// TwinCAT 3 PLC project Untitled2
// ProgramVersion: 3.1.4024.0
// libraries:
//   Tc2_MC2, * (Beckhoff Automation GmbH)
//   Tc2_NC, * (Beckhoff Automation GmbH)
//   Tc2_Standard, * (Beckhoff Automation GmbH)
//   Tc2_System, * (Beckhoff Automation GmbH)
//   Tc3_MC2_AdvancedHoming, * (Beckhoff Automation GmbH)
//   Tc3_Module, * (Beckhoff Automation GmbH)
// project tree:
//   DUTs/ ST_HandoffCmd.TcDUT, ST_HandoffStatus.TcDUT, ST_AxisPlannedReturnCmd.TcDUT, state.TcDUT
//   POUs/ Handoff.TcPOU, ArmCartesian.TcPOU, ArmCartJog.TcPOU, ArmCartJogGen.TcPOU, err.TcPOU, ArmManual.TcPOU, Axis2Sync.TcPOU, handle.TcPOU, InjectorManual.TcPOU, clear_err.TcPOU, init.TcPOU, MAIN.TcPOU, reset.TcPOU, SelfCheck.TcPOU
//   GVLs/ G.TcGVL
//   / PlcTask.TcTTO
// real-time tasks:
//   TASK PlcTask: cycle T#1ms, priority 20, ADS port 350
// motion (NC):
//   TASK NC-Task 1 SAF: cycle T#1ms, priority 4, ADS port 501
//   TASK 1: cycle T#5ms, priority 8, ADS port 511
//   AXIS Axis 1 (id 1)
//     Dynamic: Acceleration=30.3, Deceleration=30.3, Jerk=3060.3
//     Velo: SlowManual=10, FastManual=50, Maximum=30
//     OtherSettings: AllowMotionCmdToSlave=true
//     encoder EncType=19
//       EncPara: ScaleFactorNumerator=2.5, ScaleFactorDenominator=131072, Offset=230, MaxCount=#xffffffff
//     drive DrvType=16
//       DrvPara: MaxCount=#xffffffff, DriveControlDWord=#x00020100
//         Analog: TorqueSetpointScale=10, ScaleFactorActTorque=0.1
//         TimeComp: TaskDelayCycles=1
//     controller CtrType=1
//       CtrPara: PriorControlFactor=1
//         PosDiffControl: Enable=false
//         Observer: BandWidth=20
//   AXIS Axis 2 (id 2)
//     General: UnitName=°
//     Dynamic: Acceleration=10100, Deceleration=10100, Jerk=5100500
//     Velo: SlowManual=1, FastManual=5
//     OtherSettings: AllowMotionCmdToSlave=true
//     encoder EncType=19
//       EncPara: ScaleFactorNumerator=360, ScaleFactorDenominator=131072, Offset=196.397, MaxCount=#xffffffff
//     drive DrvType=16
//       DrvPara: MaxCount=#xffffffff, DriveControlDWord=#x00020000
//         Analog: TorqueSetpointScale=10, ScaleFactorActTorque=0.1
//         TimeComp: TaskDelayCycles=1
//     controller CtrType=1
//       CtrPara: PriorControlFactor=1
//         PosDiffControl: Enable=false
//         Observer: BandWidth=20
//   AXIS Axis 3 (id 3)
//     General: UnitName=°
//     Velo: SlowManual=3, FastManual=10
//     OtherSettings: AllowMotionCmdToSlave=true
//     encoder EncType=19
//       EncPara: ScaleFactorNumerator=360, ScaleFactorDenominator=131072, Offset=480, MaxCount=#xffffffff
//     drive DrvType=16
//       DrvPara: MaxCount=#xffffffff, DriveControlDWord=#x00020000
//         Analog: TorqueSetpointScale=10, ScaleFactorActTorque=0.1
//         TimeComp: TaskDelayCycles=1
//     controller CtrType=1
//       CtrPara: PriorControlFactor=1
//         PosDiffControl: Enable=false
//         Observer: BandWidth=20
//   AXIS Axis 4 (id 4)
//     General: UnitName=°
//     Dynamic: Acceleration=1570, Deceleration=1570, Jerk=2162.19
//     Velo: SlowManual=3, FastManual=10
//     OtherSettings: AllowMotionCmdToSlave=true
//     encoder EncType=19
//       EncPara: ScaleFactorNumerator=360, ScaleFactorDenominator=131072, Offset=54, MaxCount=#xffffffff
//     drive DrvType=16
//       DrvPara: MaxCount=#xffffffff, DriveControlDWord=#x00020000
//         Analog: TorqueSetpointScale=10, ScaleFactorActTorque=0.1
//         TimeComp: TaskDelayCycles=1
//     controller CtrType=1
//       CtrPara: PriorControlFactor=1
//         PosDiffControl: Enable=false
//         Observer: BandWidth=20
//   AXIS Axis 5 (id 5)
//     General: UnitName=°
//     Velo: SlowManual=3, FastManual=10
//     OtherSettings: AllowMotionCmdToSlave=true
//     encoder EncType=19
//       EncPara: ScaleFactorNumerator=360, ScaleFactorDenominator=131072, MaxCount=#xffffffff
//     drive DrvType=16
//       DrvPara: MaxCount=#xffffffff, DriveControlDWord=#x00020000
//         Analog: TorqueSetpointScale=10, ScaleFactorActTorque=0.1
//         TimeComp: TaskDelayCycles=1
//     controller CtrType=1
//       CtrPara: PriorControlFactor=1
//         Observer: BandWidth=20
//   AXIS Axis 6 (id 6)
//     Velo: SlowManual=3, FastManual=10
//     OtherSettings: AllowMotionCmdToSlave=true
//     encoder EncType=19
//       EncPara: ScaleFactorNumerator=65.94, ScaleFactorDenominator=425164.8, MaxCount=#xffffffff
//     drive DrvType=16
//       DrvPara: MaxCount=#xffffffff, DriveControlDWord=#x00020100
//         Analog: TorqueSetpointScale=10, ScaleFactorActTorque=0.1
//         TimeComp: TaskDelayCycles=1
//     controller CtrType=1
//       CtrPara: PriorControlFactor=1
//         PosDiffControl: Enable=false
//         Observer: BandWidth=20
//   AXIS Axis 7 (id 7)
//     Velo: SlowManual=3, FastManual=10
//     OtherSettings: AllowMotionCmdToSlave=true
//     encoder EncType=19
//       EncPara: ScaleFactorNumerator=360, ScaleFactorDenominator=768300, MaxCount=#xffffffff
//     drive DrvType=16
//       DrvPara: MaxCount=#xffffffff, DriveControlDWord=#x00020000
//         Analog: TorqueSetpointScale=10, ScaleFactorActTorque=0.1
//         TimeComp: TaskDelayCycles=1
//     controller CtrType=1
//       CtrPara: PriorControlFactor=1
//         PosDiffControl: Enable=false
//         Observer: BandWidth=20
//   AXIS Axis 8 (id 8)
//     Velo: SlowManual=3, FastManual=10
//     OtherSettings: AllowMotionCmdToSlave=true
//     encoder EncType=19
//       EncPara: ScaleFactorNumerator=65.94, ScaleFactorDenominator=425164.8, MaxCount=#xffffffff
//     drive DrvType=16
//       DrvPara: MaxCount=#xffffffff, DriveControlDWord=#x00020100
//         Analog: TorqueSetpointScale=10, ScaleFactorActTorque=0.1
//         TimeComp: TaskDelayCycles=1
//     controller CtrType=1
//       CtrPara: PriorControlFactor=1
//         PosDiffControl: Enable=false
//         Observer: BandWidth=20
//   AXIS Axis 9 (id 9)
//     Dynamic: Acceleration=1010, Deceleration=1010, Jerk=51005
//     Velo: SlowManual=3, FastManual=10
//     OtherSettings: AllowMotionCmdToSlave=true
//     encoder EncType=19
//       EncPara: ScaleFactorNumerator=360, ScaleFactorDenominator=758988.8, MaxCount=#xffffffff
//     drive DrvType=16
//       DrvPara: MaxCount=#xffffffff, DriveControlDWord=#x00020000
//         Analog: TorqueSetpointScale=10, ScaleFactorActTorque=0.1
//         TimeComp: TaskDelayCycles=1
//     controller CtrType=1
//       CtrPara: PriorControlFactor=1
//         Observer: BandWidth=20
//   AXIS Axis 10 (id 10)
//     Dynamic: Acceleration=2000, Deceleration=2000, Jerk=2000
//     Velo: SlowManual=3, FastManual=10
//     OtherSettings: AllowMotionCmdToSlave=true
//     encoder EncType=19
//       EncPara: ScaleFactorNumerator=65.94, ScaleFactorDenominator=425164.8, MaxCount=#xffffffff
//     drive DrvType=16
//       DrvPara: MaxCount=#xffffffff, DriveControlDWord=#x00020100
//         Analog: TorqueSetpointScale=10, ScaleFactorActTorque=0.1
//         TimeComp: TaskDelayCycles=1
//     controller CtrType=1
//       CtrPara: PriorControlFactor=1
//         PosDiffControl: Enable=false
//         Observer: BandWidth=20
//   AXIS Axis 11 (id 11)
//     Dynamic: Acceleration=375, Deceleration=375, Jerk=5625
//     Velo: SlowManual=3, FastManual=10
//     OtherSettings: AllowMotionCmdToSlave=true
//     encoder EncType=19
//       EncPara: ScaleFactorNumerator=65.94, ScaleFactorDenominator=425164.8, Inverse=true, MaxCount=#xffffffff
//     drive DrvType=16
//       DrvPara: Inverse=true, MaxCount=#xffffffff, DriveControlDWord=#x00020100
//         Analog: TorqueSetpointScale=10, ScaleFactorActTorque=0.1
//         TimeComp: TaskDelayCycles=1
//     controller CtrType=1
//       CtrPara: PriorControlFactor=1
//         PosDiffControl: Enable=false
//         Observer: BandWidth=20
//   AXIS Axis 12 (id 12)
//     Velo: SlowManual=3, FastManual=10
//     OtherSettings: AllowMotionCmdToSlave=true
//     encoder EncType=19
//       EncPara: ScaleFactorNumerator=360, ScaleFactorDenominator=768300, MaxCount=#xffffffff
//     drive DrvType=16
//       DrvPara: MaxCount=#xffffffff, DriveControlDWord=#x00020000
//         Analog: TorqueSetpointScale=10, ScaleFactorActTorque=0.1
//         TimeComp: TaskDelayCycles=1
//     controller CtrType=1
//       CtrPara: PriorControlFactor=1
//         PosDiffControl: Enable=false
//         Observer: BandWidth=20
//   AXIS Axis 13 (id 13)
//     General: UnitName=°
//     Dynamic: Acceleration=10600, Deceleration=10600, Jerk=936333
//     OtherSettings: AllowMotionCmdToSlave=true
//     encoder EncType=19
//       EncPara: ScaleFactorNumerator=360, ScaleFactorDenominator=180224, MaxCount=#xffffffff
//     drive DrvType=16
//       DrvPara: MaxCount=#xffffffff, DriveControlDWord=#x00020100
//         Analog: TorqueSetpointScale=10, ScaleFactorActTorque=0.1
//         TimeComp: TaskDelayCycles=1
//     controller CtrType=1
//       CtrPara: PriorControlFactor=1
//         PosDiffControl: Enable=false
//         Observer: BandWidth=20
//   AXIS Axis 14 (id 14)
//     General: UnitName=°
//     Dynamic: Acceleration=10400, Deceleration=10400, Jerk=1352000
//     OtherSettings: AllowMotionCmdToSlave=true
//     encoder EncType=19
//       EncPara: ScaleFactorNumerator=360, ScaleFactorDenominator=180224, MaxCount=#xffffffff
//     drive DrvType=16
//       DrvPara: MaxCount=#xffffffff, DriveControlDWord=#x00020100
//         Analog: TorqueSetpointScale=10, ScaleFactorActTorque=0.1
//         TimeComp: TaskDelayCycles=1
//     controller CtrType=1
//       CtrPara: PriorControlFactor=1
//         PosDiffControl: Enable=false
//         Observer: BandWidth=20
//   AXIS Axis 15 (id 15)
//     General: UnitName=°
//     Dynamic: Acceleration=11000, Deceleration=11000, Jerk=605000
//     OtherSettings: AllowMotionCmdToSlave=true
//     encoder EncType=19
//       EncPara: ScaleFactorNumerator=360, ScaleFactorDenominator=757760, MaxCount=#xffffffff
//     drive DrvType=16
//       DrvPara: MaxCount=#xffffffff, DriveControlDWord=#x00020100
//         Analog: TorqueSetpointScale=10, ScaleFactorActTorque=0.1
//         TimeComp: TaskDelayCycles=1
//     controller CtrType=1
//       CtrPara: PriorControlFactor=1
//         PosDiffControl: Enable=false
//         Observer: BandWidth=20
// I/O:
//   DEVICE Device 5 (EtherCAT), AmsNetId 169.254.119.135.6.1
//     Box 1 (EtherCat-control-node) [EtherCat-control-V1.6]
//     Drive 2 (Micro 4804 MZ-CAT-STO ) [Micro 4804 MZ-CAT-STO]
//     Drive 3 (TK Drive ) [EtherCAT Drive Rev:0x00010420]
//     Drive 4 (TK Drive ) [EtherCAT Drive Rev:0x00010420]
//     Drive 5 (TK Drive ) [EtherCAT Drive Rev:0x00010420]
//     Drive 6 (TK Drive ) [EtherCAT Drive Rev:0x00010420]
//     Box 7 (EtherCat-control-node) [EtherCat-control-V1.6]
//     Box 8 (EtherCat-control-node) [EtherCat-control-V1.6]
//     Drive 9 (Micro 4804 MZ-CAT-STO ) [Micro 4804 MZ-CAT-STO]
//     Drive 10 (DEN-XCR-E) [DEN-XCR-E]
//     Drive 11 (Micro 4804 MZ-CAT-STO ) [Micro 4804 MZ-CAT-STO]
//     Drive 12 (DEN-XCR-E) [DEN-XCR-E]
//     Drive 13 (Micro 4804 MZ-CAT-STO ) [Micro 4804 MZ-CAT-STO]
//     Drive 14 (Micro 4804 MZ-CAT-STO ) [Micro 4804 MZ-CAT-STO]
//     Drive 15 (CAP-XCR-E) [CAP-XCR-E]
//     Drive 16 (Micro 4804 MZ-CAT-STO ) [Micro 4804 MZ-CAT-STO]
//     Drive 17 (Micro 4804 MZ-CAT-STO ) [Micro 4804 MZ-CAT-STO]
//     Drive 18 (Micro 4804 MZ-CAT-STO ) [Micro 4804 MZ-CAT-STO]
// variable links:
//   NC-Task 1 SAF/Axes/Axis 1 <-> Device 5 (EtherCAT)/Drive 2 (Micro 4804 MZ-CAT-STO )
//     Drive/Inputs/In/nDataIn1 <-> Transmit PDO 2 mapping parameters/Following error actual value
//     Drive/Inputs/In/nDataIn3[0] <-> Transmit PDO 1 mapping parameters/Torque (current) actual value
//     Drive/Inputs/In/nDcOutputTime <-> InfoData/DcOutputShift
//     Drive/Inputs/In/nState1 <-> Transmit PDO 1 mapping parameters/Statusword
//     Drive/Inputs/In/nState2 <-> Transmit PDO 1 mapping parameters/Statusword @bit 8
//     Drive/Inputs/In/nState4 @bit 1 <-> WcState/InputToggle
//     Drive/Inputs/In/nState4 <-> WcState/WcState
//     Drive/Inputs/In/nState5 <-> Transmit PDO 4 mapping parameters/Modes of operation display
//     Drive/Outputs/Out/nCtrl1 <-> Receive PDO 1 mapping parameters/Controlword
//     Drive/Outputs/Out/nCtrl2 <-> Receive PDO 1 mapping parameters/Controlword @bit 8
//     Drive/Outputs/Out/nCtrl5 <-> Receive PDO 3 mapping parameters/Modes of operation
//     Drive/Outputs/Out/nDataOut1 <-> Receive PDO 1 mapping parameters/Target position
//     Drive/Outputs/Out/nDataOut4[0] <-> Receive PDO 3 mapping parameters/Target torque
//     Enc/Inputs/In/nDataIn1 <-> Transmit PDO 1 mapping parameters/Position actual value
//     Enc/Inputs/In/nDataIn7 <-> Transmit PDO 3 mapping parameters/Velocity actual value
//     Enc/Inputs/In/nDcInputTime <-> InfoData/DcInputShift
//     Enc/Inputs/In/nState4 @bit 1 <-> WcState/InputToggle
//     Enc/Inputs/In/nState4 <-> WcState/WcState
//   NC-Task 1 SAF/Axes/Axis 10 <-> Device 5 (EtherCAT)/Drive 13 (Micro 4804 MZ-CAT-STO )
//     Drive/Inputs/In/nDataIn1 <-> Transmit PDO 2 mapping parameters/Following error actual value
//     Drive/Inputs/In/nDataIn3[0] <-> Transmit PDO 1 mapping parameters/Torque (current) actual value
//     Drive/Inputs/In/nDcOutputTime <-> InfoData/DcOutputShift
//     Drive/Inputs/In/nState1 <-> Transmit PDO 1 mapping parameters/Statusword
//     Drive/Inputs/In/nState2 <-> Transmit PDO 1 mapping parameters/Statusword @bit 8
//     Drive/Inputs/In/nState4 @bit 1 <-> WcState/InputToggle
//     Drive/Inputs/In/nState4 <-> WcState/WcState
//     Drive/Outputs/Out/nCtrl1 <-> Receive PDO 1 mapping parameters/Controlword
//     Drive/Outputs/Out/nCtrl2 <-> Receive PDO 1 mapping parameters/Controlword @bit 8
//     Drive/Outputs/Out/nDataOut1 <-> Receive PDO 1 mapping parameters/Target position
//     Enc/Inputs/In/nDataIn1 <-> Transmit PDO 1 mapping parameters/Position actual value
//     Enc/Inputs/In/nDcInputTime <-> InfoData/DcInputShift
//     Enc/Inputs/In/nState4 @bit 1 <-> WcState/InputToggle
//     Enc/Inputs/In/nState4 <-> WcState/WcState
//   NC-Task 1 SAF/Axes/Axis 11 <-> Device 5 (EtherCAT)/Drive 14 (Micro 4804 MZ-CAT-STO )
//     Drive/Inputs/In/nDataIn1 <-> Transmit PDO 2 mapping parameters/Following error actual value
//     Drive/Inputs/In/nDataIn3[0] <-> Transmit PDO 1 mapping parameters/Torque (current) actual value
//     Drive/Inputs/In/nDcOutputTime <-> InfoData/DcOutputShift
//     Drive/Inputs/In/nState1 <-> Transmit PDO 1 mapping parameters/Statusword
//     Drive/Inputs/In/nState2 <-> Transmit PDO 1 mapping parameters/Statusword @bit 8
//     Drive/Inputs/In/nState4 @bit 1 <-> WcState/InputToggle
//     Drive/Inputs/In/nState4 <-> WcState/WcState
//     Drive/Outputs/Out/nCtrl1 <-> Receive PDO 1 mapping parameters/Controlword
//     Drive/Outputs/Out/nCtrl2 <-> Receive PDO 1 mapping parameters/Controlword @bit 8
//     Drive/Outputs/Out/nDataOut1 <-> Receive PDO 1 mapping parameters/Target position
//     Enc/Inputs/In/nDataIn1 <-> Transmit PDO 1 mapping parameters/Position actual value
//     Enc/Inputs/In/nDcInputTime <-> InfoData/DcInputShift
//     Enc/Inputs/In/nState4 @bit 1 <-> WcState/InputToggle
//     Enc/Inputs/In/nState4 <-> WcState/WcState
//   NC-Task 1 SAF/Axes/Axis 12 <-> Device 5 (EtherCAT)/Drive 15 (CAP-XCR-E)
//     Drive/Inputs/In/nState1 <-> TPDO 1 mapping parameter/Status Word
//     Drive/Inputs/In/nState2 <-> TPDO 1 mapping parameter/Status Word @bit 8
//     Drive/Inputs/In/nState4 @bit 1 <-> WcState/InputToggle
//     Drive/Inputs/In/nState4 <-> WcState/WcState
//     Drive/Inputs/In/nState5 <-> TPDO 1 mapping parameter/Operation mode display
//     Drive/Outputs/Out/nCtrl1 <-> RPDO 1 mapping parameter/Control Word
//     Drive/Outputs/Out/nCtrl2 <-> RPDO 1 mapping parameter/Control Word @bit 8
//     Drive/Outputs/Out/nCtrl5 <-> RPDO 1 mapping parameter/Operation mode
//     Drive/Outputs/Out/nDataOut1 <-> RPDO 1 mapping parameter/Position set-point
//     Drive/Outputs/Out/nDataOut2 <-> RPDO 1 mapping parameter/Velocity set-point
//     Enc/Inputs/In/nDataIn1 <-> TPDO 1 mapping parameter/Actual position
//     Enc/Inputs/In/nDataIn7 <-> TPDO 1 mapping parameter/Actual velocity
//     Enc/Inputs/In/nState4 @bit 1 <-> WcState/InputToggle
//     Enc/Inputs/In/nState4 <-> WcState/WcState
//   NC-Task 1 SAF/Axes/Axis 13 <-> Device 5 (EtherCAT)/Drive 16 (Micro 4804 MZ-CAT-STO )
//     Drive/Inputs/In/nDataIn1 <-> Transmit PDO 2 mapping parameters/Following error actual value
//     Drive/Inputs/In/nDataIn3[0] <-> Transmit PDO 1 mapping parameters/Torque (current) actual value
//     Drive/Inputs/In/nDcOutputTime <-> InfoData/DcOutputShift
//     Drive/Inputs/In/nState1 <-> Transmit PDO 1 mapping parameters/Statusword
//     Drive/Inputs/In/nState2 <-> Transmit PDO 1 mapping parameters/Statusword @bit 8
//     Drive/Inputs/In/nState4 @bit 1 <-> WcState/InputToggle
//     Drive/Inputs/In/nState4 <-> WcState/WcState
//     Drive/Outputs/Out/nCtrl1 <-> Receive PDO 1 mapping parameters/Controlword
//     Drive/Outputs/Out/nCtrl2 <-> Receive PDO 1 mapping parameters/Controlword @bit 8
//     Drive/Outputs/Out/nDataOut1 <-> Receive PDO 1 mapping parameters/Target position
//     Enc/Inputs/In/nDataIn1 <-> Transmit PDO 1 mapping parameters/Position actual value
//     Enc/Inputs/In/nDcInputTime <-> InfoData/DcInputShift
//     Enc/Inputs/In/nState4 @bit 1 <-> WcState/InputToggle
//     Enc/Inputs/In/nState4 <-> WcState/WcState
//   NC-Task 1 SAF/Axes/Axis 14 <-> Device 5 (EtherCAT)/Drive 17 (Micro 4804 MZ-CAT-STO )
//     Drive/Inputs/In/nDataIn1 <-> Transmit PDO 2 mapping parameters/Following error actual value
//     Drive/Inputs/In/nDataIn3[0] <-> Transmit PDO 1 mapping parameters/Torque (current) actual value
//     Drive/Inputs/In/nDcOutputTime <-> InfoData/DcOutputShift
//     Drive/Inputs/In/nState1 <-> Transmit PDO 1 mapping parameters/Statusword
//     Drive/Inputs/In/nState2 <-> Transmit PDO 1 mapping parameters/Statusword @bit 8
//     Drive/Inputs/In/nState4 @bit 1 <-> WcState/InputToggle
//     Drive/Inputs/In/nState4 <-> WcState/WcState
//     Drive/Outputs/Out/nCtrl1 <-> Receive PDO 1 mapping parameters/Controlword
//     Drive/Outputs/Out/nCtrl2 <-> Receive PDO 1 mapping parameters/Controlword @bit 8
//     Drive/Outputs/Out/nDataOut1 <-> Receive PDO 1 mapping parameters/Target position
//     Enc/Inputs/In/nDataIn1 <-> Transmit PDO 1 mapping parameters/Position actual value
//     Enc/Inputs/In/nDcInputTime <-> InfoData/DcInputShift
//     Enc/Inputs/In/nState4 @bit 1 <-> WcState/InputToggle
//     Enc/Inputs/In/nState4 <-> WcState/WcState
//   NC-Task 1 SAF/Axes/Axis 15 <-> Device 5 (EtherCAT)/Drive 18 (Micro 4804 MZ-CAT-STO )
//     Drive/Inputs/In/nDataIn1 <-> Transmit PDO 2 mapping parameters/Following error actual value
//     Drive/Inputs/In/nDataIn3[0] <-> Transmit PDO 1 mapping parameters/Torque (current) actual value
//     Drive/Inputs/In/nDcOutputTime <-> InfoData/DcOutputShift
//     Drive/Inputs/In/nState1 <-> Transmit PDO 1 mapping parameters/Statusword
//     Drive/Inputs/In/nState2 <-> Transmit PDO 1 mapping parameters/Statusword @bit 8
//     Drive/Inputs/In/nState4 @bit 1 <-> WcState/InputToggle
//     Drive/Inputs/In/nState4 <-> WcState/WcState
//     Drive/Outputs/Out/nCtrl1 <-> Receive PDO 1 mapping parameters/Controlword
//     Drive/Outputs/Out/nCtrl2 <-> Receive PDO 1 mapping parameters/Controlword @bit 8
//     Drive/Outputs/Out/nDataOut1 <-> Receive PDO 1 mapping parameters/Target position
//     Enc/Inputs/In/nDataIn1 <-> Transmit PDO 1 mapping parameters/Position actual value
//     Enc/Inputs/In/nDcInputTime <-> InfoData/DcInputShift
//     Enc/Inputs/In/nState4 @bit 1 <-> WcState/InputToggle
//     Enc/Inputs/In/nState4 <-> WcState/WcState
//   NC-Task 1 SAF/Axes/Axis 2 <-> Device 5 (EtherCAT)/Drive 3 (TK Drive )
//     Drive/Inputs/In/nDcOutputTime <-> InfoData/DcOutputShift
//     Drive/Inputs/In/nState1 <-> Inputs/Status word
//     Drive/Inputs/In/nState2 <-> Inputs/Status word @bit 8
//     Drive/Inputs/In/nState4 @bit 1 <-> WcState/InputToggle
//     Drive/Inputs/In/nState4 <-> WcState/WcState
//     Drive/Outputs/Out/nCtrl1 <-> Outputs/Control word
//     Drive/Outputs/Out/nCtrl2 <-> Outputs/Control word @bit 8
//     Drive/Outputs/Out/nDataOut1 <-> Outputs/Target Position
//     Enc/Inputs/In/nDataIn1 <-> Inputs/Position actual value
//     Enc/Inputs/In/nDcInputTime <-> InfoData/DcInputShift
//     Enc/Inputs/In/nState4 @bit 1 <-> WcState/InputToggle
//     Enc/Inputs/In/nState4 <-> WcState/WcState
//   NC-Task 1 SAF/Axes/Axis 3 <-> Device 5 (EtherCAT)/Drive 4 (TK Drive )
//     Drive/Inputs/In/nDcOutputTime <-> InfoData/DcOutputShift
//     Drive/Inputs/In/nState1 <-> Inputs/Status word
//     Drive/Inputs/In/nState2 <-> Inputs/Status word @bit 8
//     Drive/Inputs/In/nState4 @bit 1 <-> WcState/InputToggle
//     Drive/Inputs/In/nState4 <-> WcState/WcState
//     Drive/Outputs/Out/nCtrl1 <-> Outputs/Control word
//     Drive/Outputs/Out/nCtrl2 <-> Outputs/Control word @bit 8
//     Drive/Outputs/Out/nDataOut1 <-> Outputs/Target Position
//     Enc/Inputs/In/nDataIn1 <-> Inputs/Position actual value
//     Enc/Inputs/In/nDcInputTime <-> InfoData/DcInputShift
//     Enc/Inputs/In/nState4 @bit 1 <-> WcState/InputToggle
//     Enc/Inputs/In/nState4 <-> WcState/WcState
//   NC-Task 1 SAF/Axes/Axis 4 <-> Device 5 (EtherCAT)/Drive 5 (TK Drive )
//     Drive/Inputs/In/nDcOutputTime <-> InfoData/DcOutputShift
//     Drive/Inputs/In/nState1 <-> Inputs/Status word
//     Drive/Inputs/In/nState2 <-> Inputs/Status word @bit 8
//     Drive/Inputs/In/nState4 @bit 1 <-> WcState/InputToggle
//     Drive/Inputs/In/nState4 <-> WcState/WcState
//     Drive/Outputs/Out/nCtrl1 <-> Outputs/Control word
//     Drive/Outputs/Out/nCtrl2 <-> Outputs/Control word @bit 8
//     Drive/Outputs/Out/nDataOut1 <-> Outputs/Target Position
//     Enc/Inputs/In/nDataIn1 <-> Inputs/Position actual value
//     Enc/Inputs/In/nDcInputTime <-> InfoData/DcInputShift
//     Enc/Inputs/In/nState4 @bit 1 <-> WcState/InputToggle
//     Enc/Inputs/In/nState4 <-> WcState/WcState
//   NC-Task 1 SAF/Axes/Axis 5 <-> Device 5 (EtherCAT)/Drive 6 (TK Drive )
//     Drive/Inputs/In/nDcOutputTime <-> InfoData/DcOutputShift
//     Drive/Inputs/In/nState1 <-> Inputs/Status word
//     Drive/Inputs/In/nState2 <-> Inputs/Status word @bit 8
//     Drive/Inputs/In/nState4 @bit 1 <-> WcState/InputToggle
//     Drive/Inputs/In/nState4 <-> WcState/WcState
//     Drive/Outputs/Out/nCtrl1 <-> Outputs/Control word
//     Drive/Outputs/Out/nCtrl2 <-> Outputs/Control word @bit 8
//     Drive/Outputs/Out/nDataOut1 <-> Outputs/Target Position
//     Enc/Inputs/In/nDataIn1 <-> Inputs/Position actual value
//     Enc/Inputs/In/nDcInputTime <-> InfoData/DcInputShift
//     Enc/Inputs/In/nState4 @bit 1 <-> WcState/InputToggle
//     Enc/Inputs/In/nState4 <-> WcState/WcState
//   NC-Task 1 SAF/Axes/Axis 6 <-> Device 5 (EtherCAT)/Drive 9 (Micro 4804 MZ-CAT-STO )
//     Drive/Inputs/In/nDataIn1 <-> Transmit PDO 2 mapping parameters/Following error actual value
//     Drive/Inputs/In/nDataIn3[0] <-> Transmit PDO 1 mapping parameters/Torque (current) actual value
//     Drive/Inputs/In/nDcOutputTime <-> InfoData/DcOutputShift
//     Drive/Inputs/In/nState1 <-> Transmit PDO 1 mapping parameters/Statusword
//     Drive/Inputs/In/nState2 <-> Transmit PDO 1 mapping parameters/Statusword @bit 8
//     Drive/Inputs/In/nState4 @bit 1 <-> WcState/InputToggle
//     Drive/Inputs/In/nState4 <-> WcState/WcState
//     Drive/Outputs/Out/nCtrl1 <-> Receive PDO 1 mapping parameters/Controlword
//     Drive/Outputs/Out/nCtrl2 <-> Receive PDO 1 mapping parameters/Controlword @bit 8
//     Drive/Outputs/Out/nDataOut1 <-> Receive PDO 1 mapping parameters/Target position
//     Enc/Inputs/In/nDataIn1 <-> Transmit PDO 1 mapping parameters/Position actual value
//     Enc/Inputs/In/nDcInputTime <-> InfoData/DcInputShift
//     Enc/Inputs/In/nState4 @bit 1 <-> WcState/InputToggle
//     Enc/Inputs/In/nState4 <-> WcState/WcState
//   NC-Task 1 SAF/Axes/Axis 7 <-> Device 5 (EtherCAT)/Drive 10 (DEN-XCR-E)
//     Drive/Inputs/In/nState1 <-> TPDO 1 mapping parameter/Status Word
//     Drive/Inputs/In/nState2 <-> TPDO 1 mapping parameter/Status Word @bit 8
//     Drive/Inputs/In/nState4 @bit 1 <-> WcState/InputToggle
//     Drive/Inputs/In/nState4 <-> WcState/WcState
//     Drive/Inputs/In/nState5 <-> TPDO 1 mapping parameter/Operation mode display
//     Drive/Outputs/Out/nCtrl1 <-> RPDO 1 mapping parameter/Control Word
//     Drive/Outputs/Out/nCtrl2 <-> RPDO 1 mapping parameter/Control Word @bit 8
//     Drive/Outputs/Out/nCtrl5 <-> RPDO 1 mapping parameter/Operation mode
//     Drive/Outputs/Out/nDataOut1 <-> RPDO 1 mapping parameter/Position set-point
//     Drive/Outputs/Out/nDataOut2 <-> RPDO 1 mapping parameter/Velocity set-point
//     Enc/Inputs/In/nDataIn1 <-> TPDO 1 mapping parameter/Actual position
//     Enc/Inputs/In/nDataIn7 <-> TPDO 1 mapping parameter/Actual velocity
//     Enc/Inputs/In/nState4 @bit 1 <-> WcState/InputToggle
//     Enc/Inputs/In/nState4 <-> WcState/WcState
//   NC-Task 1 SAF/Axes/Axis 8 <-> Device 5 (EtherCAT)/Drive 11 (Micro 4804 MZ-CAT-STO )
//     Drive/Inputs/In/nDataIn1 <-> Transmit PDO 2 mapping parameters/Following error actual value
//     Drive/Inputs/In/nDataIn3[0] <-> Transmit PDO 1 mapping parameters/Torque (current) actual value
//     Drive/Inputs/In/nDcOutputTime <-> InfoData/DcOutputShift
//     Drive/Inputs/In/nState1 <-> Transmit PDO 1 mapping parameters/Statusword
//     Drive/Inputs/In/nState2 <-> Transmit PDO 1 mapping parameters/Statusword @bit 8
//     Drive/Inputs/In/nState4 @bit 1 <-> WcState/InputToggle
//     Drive/Inputs/In/nState4 <-> WcState/WcState
//     Drive/Outputs/Out/nCtrl1 <-> Receive PDO 1 mapping parameters/Controlword
//     Drive/Outputs/Out/nCtrl2 <-> Receive PDO 1 mapping parameters/Controlword @bit 8
//     Drive/Outputs/Out/nDataOut1 <-> Receive PDO 1 mapping parameters/Target position
//     Enc/Inputs/In/nDataIn1 <-> Transmit PDO 1 mapping parameters/Position actual value
//     Enc/Inputs/In/nDcInputTime <-> InfoData/DcInputShift
//     Enc/Inputs/In/nState4 @bit 1 <-> WcState/InputToggle
//     Enc/Inputs/In/nState4 <-> WcState/WcState
//   NC-Task 1 SAF/Axes/Axis 9 <-> Device 5 (EtherCAT)/Drive 12 (DEN-XCR-E)
//     Drive/Inputs/In/nState1 <-> TPDO 1 mapping parameter/Status Word
//     Drive/Inputs/In/nState2 <-> TPDO 1 mapping parameter/Status Word @bit 8
//     Drive/Inputs/In/nState4 @bit 1 <-> WcState/InputToggle
//     Drive/Inputs/In/nState4 <-> WcState/WcState
//     Drive/Inputs/In/nState5 <-> TPDO 1 mapping parameter/Operation mode display
//     Drive/Outputs/Out/nCtrl1 <-> RPDO 1 mapping parameter/Control Word
//     Drive/Outputs/Out/nCtrl2 <-> RPDO 1 mapping parameter/Control Word @bit 8
//     Drive/Outputs/Out/nCtrl5 <-> RPDO 1 mapping parameter/Operation mode
//     Drive/Outputs/Out/nDataOut1 <-> RPDO 1 mapping parameter/Position set-point
//     Drive/Outputs/Out/nDataOut2 <-> RPDO 1 mapping parameter/Velocity set-point
//     Enc/Inputs/In/nDataIn1 <-> TPDO 1 mapping parameter/Actual position
//     Enc/Inputs/In/nDataIn7 <-> TPDO 1 mapping parameter/Actual velocity
//     Enc/Inputs/In/nState4 @bit 1 <-> WcState/InputToggle
//     Enc/Inputs/In/nState4 <-> WcState/WcState
//   Untitled2/Untitled2 Instance <-> Device 5 (EtherCAT)/Box 7 (EtherCat-control-node)
//     PlcTask Inputs/G.fn_2_value <-> Data Inputs/Data_4
//     PlcTask Inputs/G.ft_2_value <-> Data Inputs/Data_3
//     PlcTask Outputs/G.cylinder3_value <-> Outputs/Value_1
//     PlcTask Outputs/G.cylinder4_value <-> Outputs/Value_2
//   Untitled2/Untitled2 Instance <-> Device 5 (EtherCAT)/Box 8 (EtherCat-control-node)
//     PlcTask Inputs/G.fn_1_value <-> Data Inputs/Data_4
//     PlcTask Inputs/G.ft_1_value <-> Data Inputs/Data_3
//     PlcTask Outputs/G.cylinder1_value <-> Outputs/Value_1
//     PlcTask Outputs/G.cylinder2_value <-> Outputs/Value_2
//     PlcTask Outputs/G.cylinder5_value <-> Outputs/Value_3
//   Untitled2/Untitled2 Instance <-> NC-Task 1 SAF/Axes/Axis 1
//     PlcTask Inputs/G.arm_axis[1].NcToPlc <-> Outputs/ToPlc
//     PlcTask Outputs/G.arm_axis[1].PlcToNc <-> Inputs/FromPlc
//   Untitled2/Untitled2 Instance <-> NC-Task 1 SAF/Axes/Axis 10
//     PlcTask Inputs/G.axis[5].NcToPlc <-> Outputs/ToPlc
//     PlcTask Outputs/G.axis[5].PlcToNc <-> Inputs/FromPlc
//   Untitled2/Untitled2 Instance <-> NC-Task 1 SAF/Axes/Axis 11
//     PlcTask Inputs/G.axis[6].NcToPlc <-> Outputs/ToPlc
//     PlcTask Outputs/G.axis[6].PlcToNc <-> Inputs/FromPlc
//   Untitled2/Untitled2 Instance <-> NC-Task 1 SAF/Axes/Axis 12
//     PlcTask Inputs/G.axis[7].NcToPlc <-> Outputs/ToPlc
//     PlcTask Outputs/G.axis[7].PlcToNc <-> Inputs/FromPlc
//   Untitled2/Untitled2 Instance <-> NC-Task 1 SAF/Axes/Axis 13
//     PlcTask Inputs/G.inject_axis[1].NcToPlc <-> Outputs/ToPlc
//     PlcTask Outputs/G.inject_axis[1].PlcToNc <-> Inputs/FromPlc
//   Untitled2/Untitled2 Instance <-> NC-Task 1 SAF/Axes/Axis 14
//     PlcTask Inputs/G.inject_axis[2].NcToPlc <-> Outputs/ToPlc
//     PlcTask Outputs/G.inject_axis[2].PlcToNc <-> Inputs/FromPlc
//   Untitled2/Untitled2 Instance <-> NC-Task 1 SAF/Axes/Axis 15
//     PlcTask Inputs/G.axis2_sync_axis.NcToPlc <-> Outputs/ToPlc
//     PlcTask Outputs/G.axis2_sync_axis.PlcToNc <-> Inputs/FromPlc
//   Untitled2/Untitled2 Instance <-> NC-Task 1 SAF/Axes/Axis 2
//     PlcTask Inputs/G.arm_axis[2].NcToPlc <-> Outputs/ToPlc
//     PlcTask Outputs/G.arm_axis[2].PlcToNc <-> Inputs/FromPlc
//   Untitled2/Untitled2 Instance <-> NC-Task 1 SAF/Axes/Axis 3
//     PlcTask Inputs/G.arm_axis[3].NcToPlc <-> Outputs/ToPlc
//     PlcTask Outputs/G.arm_axis[3].PlcToNc <-> Inputs/FromPlc
//   Untitled2/Untitled2 Instance <-> NC-Task 1 SAF/Axes/Axis 4
//     PlcTask Inputs/G.arm_axis[4].NcToPlc <-> Outputs/ToPlc
//     PlcTask Outputs/G.arm_axis[4].PlcToNc <-> Inputs/FromPlc
//   Untitled2/Untitled2 Instance <-> NC-Task 1 SAF/Axes/Axis 5
//     PlcTask Inputs/G.arm_axis[5].NcToPlc <-> Outputs/ToPlc
//     PlcTask Outputs/G.arm_axis[5].PlcToNc <-> Inputs/FromPlc
//   Untitled2/Untitled2 Instance <-> NC-Task 1 SAF/Axes/Axis 6
//     PlcTask Inputs/G.axis[1].NcToPlc <-> Outputs/ToPlc
//     PlcTask Outputs/G.axis[1].PlcToNc <-> Inputs/FromPlc
//   Untitled2/Untitled2 Instance <-> NC-Task 1 SAF/Axes/Axis 7
//     PlcTask Inputs/G.axis[2].NcToPlc <-> Outputs/ToPlc
//     PlcTask Outputs/G.axis[2].PlcToNc <-> Inputs/FromPlc
//   Untitled2/Untitled2 Instance <-> NC-Task 1 SAF/Axes/Axis 8
//     PlcTask Inputs/G.axis[3].NcToPlc <-> Outputs/ToPlc
//     PlcTask Outputs/G.axis[3].PlcToNc <-> Inputs/FromPlc
//   Untitled2/Untitled2 Instance <-> NC-Task 1 SAF/Axes/Axis 9
//     PlcTask Inputs/G.axis[4].NcToPlc <-> Outputs/ToPlc
//     PlcTask Outputs/G.axis[4].PlcToNc <-> Inputs/FromPlc

CONFIGURATION Untitled2
    RESOURCE PLC ON TwinCAT3
        TASK PlcTask(INTERVAL := T#1ms, PRIORITY := 20);
        PROGRAM MAIN WITH PlcTask : MAIN;
    END_RESOURCE
END_CONFIGURATION

// ---- DUTs/ST_HandoffCmd.TcDUT
{attribute 'pack_mode' := '1'}
TYPE ST_HandoffCmd :
STRUCT
    leg_mask : BYTE;
    target_abs : ARRAY[1..2] OF LREAL;
    velocity : ARRAY[1..2] OF LREAL;
    acc : ARRAY[1..2] OF LREAL;
    dec : ARRAY[1..2] OF LREAL;
    jerk : ARRAY[1..2] OF LREAL;
    cyl_clamp : ARRAY[1..4] OF WORD;
    cyl_open : ARRAY[1..4] OF WORD;
    wait_ms : ARRAY[1..2] OF ARRAY[1..4] OF UINT;
    request_id : UDINT;
END_STRUCT
END_TYPE

// ---- DUTs/ST_HandoffStatus.TcDUT
{attribute 'pack_mode' := '1'}
TYPE ST_HandoffStatus :
STRUCT
    ack_id : UDINT;
    phase : INT;
    phase_seq : UDINT;
    done_id : UDINT;
    result : INT;
    error_code : UDINT;
    error_axis : INT;
    nc_error_code : UDINT;
    reject_reason : INT; // 1=忙，2=状态不允许，3=参数非法
    leg_mask : BYTE; // 受理腿集合，供数据端重启后接管
    phase_ms : ARRAY[1..8] OF UDINT; // 10/20/30/40/50、轴1运动、轴6运动、保留
END_STRUCT
END_TYPE

// ---- DUTs/ST_AxisPlannedReturnCmd.TcDUT
TYPE ST_AxisPlannedReturnCmd :
STRUCT
	Req			: BOOL;
	Busy		: BOOL;
	Done		: BOOL;
	Error		: BOOL;
	ErrorId		: UDINT;
	TargetAbs	: LREAL;
	Velocity	: LREAL;
	Acc			: LREAL;
	Dec			: LREAL;
	Jerk		: LREAL;
END_STRUCT
END_TYPE

// ---- DUTs/state.TcDUT
TYPE state :
(
	_init := 0,		//全下电
	_jog1,			//一二轴回零位
	_jog2,			//三轴回零
	_jog3,			//其余轴回零
	_trans,	//进入运输位
	_trans_wait,	//进入运输位
	_handle,		//跟随手柄运动
	_self_check,    //上电自检
	_clear_err,
	_err,
	_reset
)INT;

END_TYPE

// ---- GVLs/G.TcGVL
{attribute 'qualified_only'}
VAR_GLOBAL
	// 第五轮恢复诊断与寻参复用接口。
	err_backoff_active : ARRAY[1..7] OF BOOL;
	err_backoff_failed : ARRAY[1..7] OF BOOL;
	axis2_sync_error : BOOL;
	axis2_sync_error_id : UDINT;
	homing_restore_req : BOOL;
	homing_restore_leftlimit : ARRAY[1..7] OF LREAL;
	homing_restore_init_pos : ARRAY[1..7] OF LREAL;
	homing_restore_status : DINT;
	homing_restore_reject_reason : DINT;
	//专有变量
	gen_state			:	state := _init;
	axis				:	ARRAY[1..7] OF axis_REF;
	power_				:	ARRAY[1..7] OF MC_Power;
	power_output		:	ARRAY[1..7] OF ST_McOutputs;
	axis_Reset			:	ARRAY[1..7] OF MC_Reset;
	reset_output		:	ARRAY[1..7] OF ST_McOutputs;
	SetPointGenEnable	:	ARRAY[1..7] OF MC_ExtSetPointGenEnable;
	SetPointGenDisable	:	ARRAY[1..7] OF MC_ExtSetPointGenDisable;
	SetPointGenEnable_output,	SetPointGenDisable_output	: ARRAY[1..7] OF ST_McOutputs;
	move_jog			: 	ARRAY [1..7] OF MC_Jog;
	enable,	disable		:	BOOL;	//跟随运动变量
	flag:INT:=0;
	flagpos:LREAL:=0; // 遗留调试量，当前无业务读取
    //其他变量
    init_pos			: ARRAY[1..7] OF LREAL := [30, 9, 0, 0, 0, 30, 13];
    refer,Act_pos,act_h,act_hf	: ARRAY[1..7] OF LREAL;
    
	// 自检相关变量
    leftlimit           : ARRAY[1..7] OF LREAL;
	act_pos_from_left	: ARRAY[1..7] OF LREAL;
	refer_from_left		: ARRAY[1..7] OF LREAL;
    self_check_done     : BOOL := FALSE;
	selfcheck_start_req  : BOOL := FALSE;
	selfcheck_status     : DINT := 0; // 0=未就绪，1=等待启动，2=运行中，3=参数拒绝
	selfcheck_target_from_left : ARRAY[1..7] OF LREAL := [96,0,500,0,530,580,0];
	startup_loading_ready : BOOL := FALSE; // TRUE=自检刚完成且仍允许按标准器械装卸姿态启动；上位机开始控制前消费为 FALSE
	handle_reinit_req	: BOOL := FALSE;
	handle_reinit_done	: BOOL := FALSE;
	selfcheck_reset_req : BOOL := FALSE;
	selfcheck_stu		: ARRAY[1..7] OF INT;
	selfcheck_all_reach_limit : BOOL := FALSE;

	// 急停/掉使能冻结：用于通知上位机停止写 refer，并在恢复时触发重同步
	estop_hold_req		: BOOL := FALSE;

	// ADS 上位机心跳看门狗：上位机保持会话号不变并递增心跳序号。
	// 超时后必须先恢复心跳，再置 host_recover_req；PLC 停稳后清除请求并启动重初始化。
	// host_comm_timeout=FALSE 表示请求已受理，handle_reinit_done=TRUE 表示重初始化完成。
	host_session_id			: UDINT := 0;
	host_heartbeat_sequence	: UDINT := 0;
	host_recover_req		: BOOL := FALSE;
	host_comm_timeout		: BOOL := TRUE;

    handoff_cmd : ST_HandoffCmd;
    handoff_status : ST_HandoffStatus;
    handoff_takeover_id : UDINT;
    handoff_if_version : UDINT := 1;
    cyl_cmd : ARRAY[1..4] OF WORD;
	axis4_fwd_req		: BOOL := FALSE;
	axis4_rev_req		: BOOL := FALSE;
	axis4_manual_busy	: BOOL := FALSE;
	axis4_manual_done	: BOOL := FALSE;
	axis4_manual_error	: BOOL := FALSE;
	axis4_manual_error_id : UDINT := 0;


	// 速度门限与参考缓动（参考“方式10-仿真”风格）
	v_limit				: ARRAY[1..7] OF LREAL := [7.5,7.5,1.5,1.5,1.5,7.5,1.5];
	ref_slow			: ARRAY[1..7] OF LREAL := [0,0,0,0,0,0,0];

	// PID 参数（可按轴整定）及状态量
	// 以下 PID 参数已废弃：控制路径已改为速率限制+滑动平均+轨迹滤波，上位机勿依赖。
	Kp					: ARRAY[1..7] OF LREAL := [0.14,0.14,0.14,0.14,0.14,0.14,0.14];
	Ki					: ARRAY[1..7] OF LREAL := [0.016,0.016,0.016,0.016,0.016,0.016,0.016];
	Kd					: ARRAY[1..7] OF LREAL := [0.1,0.1,0.1,0.1,0.1,0.1,0.1];
	pid_i				: ARRAY[1..7] OF LREAL := [0,0,0,0,0,0,0];
	pid_e_prev			: ARRAY[1..7] OF LREAL := [0,0,0,0,0,0,0];
	pid_i_limit			: ARRAY[1..7] OF LREAL := [100,100,100,100,100,100,100];

	// ========== 定位臂 5 轴独立点动控制变量 ==========
	arm_axis			: ARRAY[1..5] OF AXIS_REF;	// 定位臂轴对象，链接到 NC Axis 1..5
	arm_manual_enable	: BOOL := FALSE;			// 定位臂手动控制总使能，FALSE 时所有点动请求无效
	arm_enable_req		: ARRAY[1..5] OF BOOL := [FALSE,FALSE,FALSE,FALSE,FALSE];	// TRUE=对应轴保持上电
	arm_reset_req		: ARRAY[1..5] OF BOOL := [FALSE,FALSE,FALSE,FALSE,FALSE];	// TRUE=请求清错，PLC 完成后自动清零
	arm_jog_pos_req		: ARRAY[1..5] OF BOOL := [FALSE,FALSE,FALSE,FALSE,FALSE];	// UI 正向点动按钮，按下 TRUE、松开 FALSE
	arm_jog_neg_req		: ARRAY[1..5] OF BOOL := [FALSE,FALSE,FALSE,FALSE,FALSE];	// UI 反向点动按钮，按下 TRUE、松开 FALSE
	arm_jog_velocity	: ARRAY[1..5] OF LREAL := [5.0,5.0,5.0,5.0,5.0];
	arm_jog_acc		: ARRAY[1..5] OF LREAL := [50.0,50.0,50.0,50.0,50.0];
	arm_jog_dec		: ARRAY[1..5] OF LREAL := [50.0,50.0,50.0,50.0,50.0];
	arm_jog_jerk		: ARRAY[1..5] OF LREAL := [500.0,500.0,500.0,500.0,500.0];
	arm_power_output	: ARRAY[1..5] OF ST_McOutputs;
	arm_reset_output	: ARRAY[1..5] OF ST_McOutputs;
	arm_act_pos		: ARRAY[1..5] OF LREAL;
	arm_act_vel		: ARRAY[1..5] OF LREAL;
	arm_motion_busy		: ARRAY[1..5] OF BOOL := [FALSE,FALSE,FALSE,FALSE,FALSE];
	arm_motion_done		: ARRAY[1..5] OF BOOL := [FALSE,FALSE,FALSE,FALSE,FALSE];
	arm_motion_error	: ARRAY[1..5] OF BOOL := [FALSE,FALSE,FALSE,FALSE,FALSE];
	arm_motion_error_id	: ARRAY[1..5] OF UDINT := [0,0,0,0,0];
	arm_cmd_dir		: ARRAY[1..5] OF SINT := [0,0,0,0,0];	// -1=反向，0=停止，1=正向
	arm_cmd_conflict	: ARRAY[1..5] OF BOOL := [FALSE,FALSE,FALSE,FALSE,FALSE];	// 正反向同时请求
	// 归零曲线接口：先写数据再递增request。
	arm_curve_data : ARRAY[0..16] OF LREAL;
	arm_curve_request : UDINT;
	arm_curve_ack : UDINT;
	arm_curve_cancel : BOOL := TRUE;
	arm_curve_heartbeat : UDINT;
	arm_curve_owned : BOOL;
	arm_curve_state : UDINT; // 0空闲，1执行，2完成，3取消，4错误
	arm_curve_error : UDINT;
	arm_curve_progress : LREAL;
	// 末端点动请求：毫米/秒或度/秒；保活计数按住期间递增。
	arm_cjog_mode : INT;
	arm_cjog_dir : INT;
	arm_cjog_speed : LREAL;
	arm_cjog_alive : UDINT;
	arm_cjog_owned : BOOL;
	arm_cjog_state : UDINT; // 0空闲，1使能，2运动，3减速，4释放
	arm_cjog_error : UDINT;
	arm_cjog_limited : BOOL;
	arm_cjog_path_speed : LREAL;
	arm_cjog_if_version : UDINT := 1;

	// ========== Axis15 同步接口 ==========
	// 独立链接到 NC Axis 15，与业务轴2（NC Axis 7）同步旋转。
	axis2_sync_axis	: AXIS_REF;

	// ========== 注射器轴控制接口 ==========
	// inject_axis[1] -> NC Axis 13 / Drive 16，inject_axis[2] -> NC Axis 14 / Drive 17。
	inject_axis		: ARRAY[1..2] OF AXIS_REF;
	inject_push_req	: ARRAY[1..2] OF BOOL := [FALSE,FALSE];
	inject_pull_req	: ARRAY[1..2] OF BOOL := [FALSE,FALSE];

	// ========== 电缸控制变量 ==========
	cylinder1_value		AT %Q* : WORD;		// 电缸1控制值 (安装在夹持机构上)
	cylinder2_value		AT %Q* : WORD;		// 电缸2控制值 (安装在轴1机构上)
	cylinder3_value		AT %Q* : WORD;		// 电缸3控制值 (安装在轴5机构上)
	cylinder4_value		AT %Q* : WORD;		// 电缸4控制值 (安装在轴6机构上)
	cylinder5_value		AT %Q* : WORD;		// 电缸5控制值 (安装在轴3机构上控制y阀)
	cylinder5_cmd		: WORD := 2000;		// 历史兼容缓存，当前正式控制不写此变量
	cylinder5_press_req	: BOOL := FALSE;	// Y阀请求（TRUE=打开，输出500；FALSE=关闭，输出2000）
	
	
	ft_1_value			AT %I* : INT;
	fn_1_value			AT %I* : INT;
	fn_2_value			AT %I* : INT;
	ft_2_value			AT %I* : INT;



	// 手柄模式最近一次急停入口快照：计数增加后读取，自动恢复不清除；数组下标为轴号。
	estop_diag_count : UDINT;
	estop_diag_host_timeout : BOOL;
	estop_diag_axis : ARRAY[1..7] OF ST_AxisStatus;
	estop_diag_power : ARRAY[1..7] OF ST_McOutputs;
	estop_diag_reset : ARRAY[1..7] OF ST_McOutputs;
	estop_diag_power_enable : ARRAY[1..7] OF BOOL;
	estop_diag_power_positive : ARRAY[1..7] OF BOOL;
	estop_diag_power_negative : ARRAY[1..7] OF BOOL;
	estop_diag_return_state : ARRAY[1..7] OF INT;
	estop_diag_return_cmd : ARRAY[1..7] OF ST_AxisPlannedReturnCmd;
	estop_diag_move_error : ARRAY[1..7] OF BOOL;
	estop_diag_move_aborted : ARRAY[1..7] OF BOOL;
	estop_diag_enable_error : ARRAY[1..7] OF BOOL;
	estop_diag_disable_error : ARRAY[1..7] OF BOOL;
	estop_diag_move_error_id : ARRAY[1..7] OF UDINT;
	estop_diag_enable_error_id : ARRAY[1..7] OF UDINT;
	estop_diag_disable_error_id : ARRAY[1..7] OF UDINT;
	estop_diag_act_pos : ARRAY[1..7] OF LREAL;
	estop_diag_act_vel : ARRAY[1..7] OF LREAL;
	estop_diag_feed_pos : ARRAY[1..7] OF LREAL;
	estop_diag_feed_vel : ARRAY[1..7] OF LREAL;
	estop_diag_refer_abs : ARRAY[1..7] OF LREAL;
END_VAR
VAR_GLOBAL CONSTANT
	rslimit_distance : ARRAY[1..7] OF LREAL := [99.0, 0.0, 666.0, 0.0, 688.0, 688.0, 0.0];
	recovery_wait_timeout : TIME := T#2S;
	recovery_max_retries : UINT := 3;
	err_backoff_distance : LREAL := 2.0;
	err_backoff_velocity : LREAL := 5.0;
	err_backoff_acc : LREAL := 50.0;
	axis15_reset_pulse : TIME := T#200MS;
	axis15_reset_interval : TIME := T#2S;
    handoff_err_rejected : UDINT := 1;
    handoff_err_disable : UDINT := 2;
    handoff_err_move : UDINT := 3;
    handoff_err_timeout : UDINT := 4;
    handoff_err_interrupted : UDINT := 5;
END_VAR

// ---- POUs/MAIN.TcPOU
PROGRAM MAIN
VAR
    handoff_called : BOOL;
	init_		:		init;
	handle1_	:		handle;
	clear_err_	:		clear_err;
	err_		:		err;
	reset_		:		reset;
	self_check_ :       SelfCheck;
	arm_manual_ :       ArmManual;
	arm_cartesian_ :    ArmCartesian;
	arm_cart_jog_ :     ArmCartJog;
	axis2_sync_ :       Axis2Sync;
	injector_manual_ :  InjectorManual;
	axis6_enable_negative : BOOL := TRUE;
	selfcheck_started : BOOL := FALSE;
	selfcheck_target_latched : ARRAY[1..7] OF LREAL;
	host_watchdog_timer : TON;
	host_last_heartbeat_sequence : UDINT;
	host_last_session_id : UDINT;
	host_session_changed : BOOL;
	host_heartbeat_changed : BOOL;
	host_heartbeat_seen : BOOL;
	i:INT;
	last_dispatched_state : state := _init;
	dispatched_state : state;
	restore_ready : BOOL;
	restore_pending : BOOL;
	restore_disabled : BOOL;
	restore_disable_error : BOOL;
END_VAR

FOR i:=1 TO 7 DO
	G.axis[i]();	
END_FOR

// 注射器 NC 轴刷新 AXIS_REF，由独立点动 POU 控制，不进入业务状态机。
FOR i:=1 TO 2 DO
	G.inject_axis[i]();
END_FOR

IF TwinCAT_SystemInfoVarList._TaskInfo[1].FirstCycle THEN
	G.gen_state := _init;
	G.self_check_done := FALSE;
	G.selfcheck_start_req := FALSE;
	G.selfcheck_status := 0;
	G.handle_reinit_req := FALSE;
	G.handle_reinit_done := FALSE;
	G.estop_hold_req := FALSE;
	G.selfcheck_reset_req := TRUE;
	FOR i:=1 TO 7 DO
		G.SetPointGenEnable[i].Execute := FALSE;
		G.SetPointGenDisable[i].Execute := FALSE;
		G.axis_Reset[i].Execute := FALSE;
	END_FOR
	G.arm_manual_enable := FALSE;
	FOR i:=1 TO 5 DO
		// PLC 启动时定位臂必须保持断使能，不能因为残留请求自动上电。
		G.arm_enable_req[i] := FALSE;
		G.arm_reset_req[i] := FALSE;
		G.arm_jog_pos_req[i] := FALSE;
		G.arm_jog_neg_req[i] := FALSE;
	END_FOR
END_IF

// ==================== 全局主机通信看门狗 (2s 超时) ====================
host_session_changed := G.host_session_id <> host_last_session_id;
host_heartbeat_changed := host_session_changed OR
	(G.host_heartbeat_sequence <> host_last_heartbeat_sequence);

IF host_session_changed THEN
	IF host_last_session_id <> 0 THEN
		G.host_comm_timeout := TRUE;
	END_IF
	host_last_session_id := G.host_session_id;
END_IF

IF host_heartbeat_changed THEN
	host_last_heartbeat_sequence := G.host_heartbeat_sequence;
END_IF

host_heartbeat_seen := G.host_session_id <> 0;
host_watchdog_timer(
	IN:=host_heartbeat_seen AND NOT host_heartbeat_changed,
	PT:=T#2S
);
IF (NOT host_heartbeat_seen) OR host_watchdog_timer.Q THEN
	G.host_comm_timeout := TRUE;
ELSIF G.gen_state <> _handle THEN
	// 自检前等待阶段：收到上位机恢复请求且心跳正常时解除超时
	IF G.host_recover_req THEN
		G.host_comm_timeout := FALSE;
		G.host_recover_req := FALSE;
	END_IF
END_IF
// ======================================================================
	
arm_manual_();
arm_cartesian_();
arm_cart_jog_();
axis2_sync_();
injector_manual_();

// 轴6自检触发左限位后只关闭负向许可，保留正向脱离限位的能力。
axis6_enable_negative := NOT ((G.gen_state = _self_check) AND G.axis[6].Status.DriveLimitActive);
POWERED();
IF G.gen_state <> _handle THEN
	SETPOSITIONGEN();
END_IF
RESETED();

IF G.gen_state <> _self_check THEN
	selfcheck_started := FALSE;
	G.selfcheck_start_req := FALSE;
	G.selfcheck_status := 0;
END_IF

dispatched_state := G.gen_state;
handoff_called := FALSE;
CASE G.gen_state OF
	_init:			init_();
	_self_check:
        IF G.homing_restore_req THEN
            G.homing_restore_req := FALSE;
            G.homing_restore_status := 0;
            G.homing_restore_reject_reason := 0;
            restore_pending := TRUE;
        END_IF
        IF restore_pending THEN
            restore_ready := NOT selfcheck_started AND NOT G.selfcheck_start_req;
            restore_disabled := TRUE;
            restore_disable_error := FALSE;
            FOR i:=1 TO 7 DO
                IF NOT G.power_output[i].Done OR G.axis[i].Status.Error OR G.axis[i].Status.DriveDeviceError
                    OR G.power_output[i].Error OR G.reset_output[i].Error THEN restore_ready := FALSE; END_IF
                G.SetPointGenEnable[i].Execute := FALSE;
                G.SetPointGenDisable[i](Axis:=G.axis[i], Execute:=TRUE);
                IF G.SetPointGenDisable[i].Error THEN restore_disable_error := TRUE; END_IF
                IF NOT (G.SetPointGenDisable[i].Done OR NOT G.SetPointGenDisable[i].Enabled) THEN restore_disabled := FALSE; END_IF
            END_FOR
            IF NOT restore_ready OR restore_disable_error THEN
                restore_pending := FALSE;
                G.homing_restore_status := 2;
                IF restore_disable_error THEN G.homing_restore_reject_reason := 2;
                ELSE G.homing_restore_reject_reason := 1; END_IF
                FOR i:=1 TO 7 DO G.SetPointGenDisable[i].Execute := FALSE; END_FOR
            ELSE
			IF restore_disabled THEN
				G.leftlimit := G.homing_restore_leftlimit;
				G.init_pos := G.homing_restore_init_pos;
				G.cylinder1_value := 1000;
				G.cylinder2_value := 150;
				G.cylinder3_value := 1000;
				G.cylinder4_value := 150;
				G.self_check_done := TRUE;
				G.startup_loading_ready := FALSE;
				G.handle_reinit_req := TRUE;
				FOR i:=1 TO 7 DO
					G.SetPointGenDisable[i](Axis:=G.axis[i], Execute:=FALSE);
					G.Act_pos[i] := G.axis[i].NcToPlc.ActPos - G.init_pos[i];
					G.act_pos_from_left[i] := G.axis[i].NcToPlc.ActPos - G.leftlimit[i];
					G.refer[i] := G.Act_pos[i];
					G.ref_slow[i] := G.Act_pos[i];
					G.act_h[i] := G.Act_pos[i];
					G.act_hf[i] := G.Act_pos[i];
					G.refer_from_left[i] := G.act_pos_from_left[i];
				END_FOR
				G.homing_restore_status := 1;
				G.homing_restore_reject_reason := 0;
				G.gen_state := _handle;
				restore_pending := FALSE;
                END_IF
            END_IF
        END_IF
		IF (G.gen_state = _self_check) AND NOT selfcheck_started AND NOT restore_pending THEN
			IF G.selfcheck_status <> 3 THEN G.selfcheck_status := 1; END_IF
			IF G.selfcheck_start_req THEN
				G.selfcheck_start_req := FALSE;
				IF G.selfcheck_target_from_left[1] >= 5.0 AND G.selfcheck_target_from_left[1] <= 96.0
					AND G.selfcheck_target_from_left[3] >= 10.0 AND G.selfcheck_target_from_left[3] <= 650.0
					AND G.selfcheck_target_from_left[5] >= 10.0 AND G.selfcheck_target_from_left[5] <= 670.0
					AND G.selfcheck_target_from_left[6] >= 10.0 AND G.selfcheck_target_from_left[6] <= 670.0
					AND G.selfcheck_target_from_left[1] <= G.selfcheck_target_from_left[3]
					AND G.selfcheck_target_from_left[3] <= G.selfcheck_target_from_left[5]
					AND G.selfcheck_target_from_left[5] <= G.selfcheck_target_from_left[6] THEN
					selfcheck_target_latched := G.selfcheck_target_from_left;
					selfcheck_started := TRUE;
					G.selfcheck_status := 2;
				ELSE
					G.selfcheck_status := 3;
				END_IF
			END_IF
		END_IF
		IF selfcheck_started THEN
			self_check_(init_target_from_left := selfcheck_target_latched);
		END_IF
	_handle:		handoff_called := TRUE; handle1_();	
		SETPOSITIONGEN();
	_clear_err:		clear_err_();	
	_err:			err_(enter := last_dispatched_state <> _err);
	_reset:			reset_();
END_CASE
IF NOT handoff_called THEN
    handle1_.handoff(ready:=FALSE, interrupted:=TRUE);
END_IF
last_dispatched_state := dispatched_state;

ACTION POWERED:
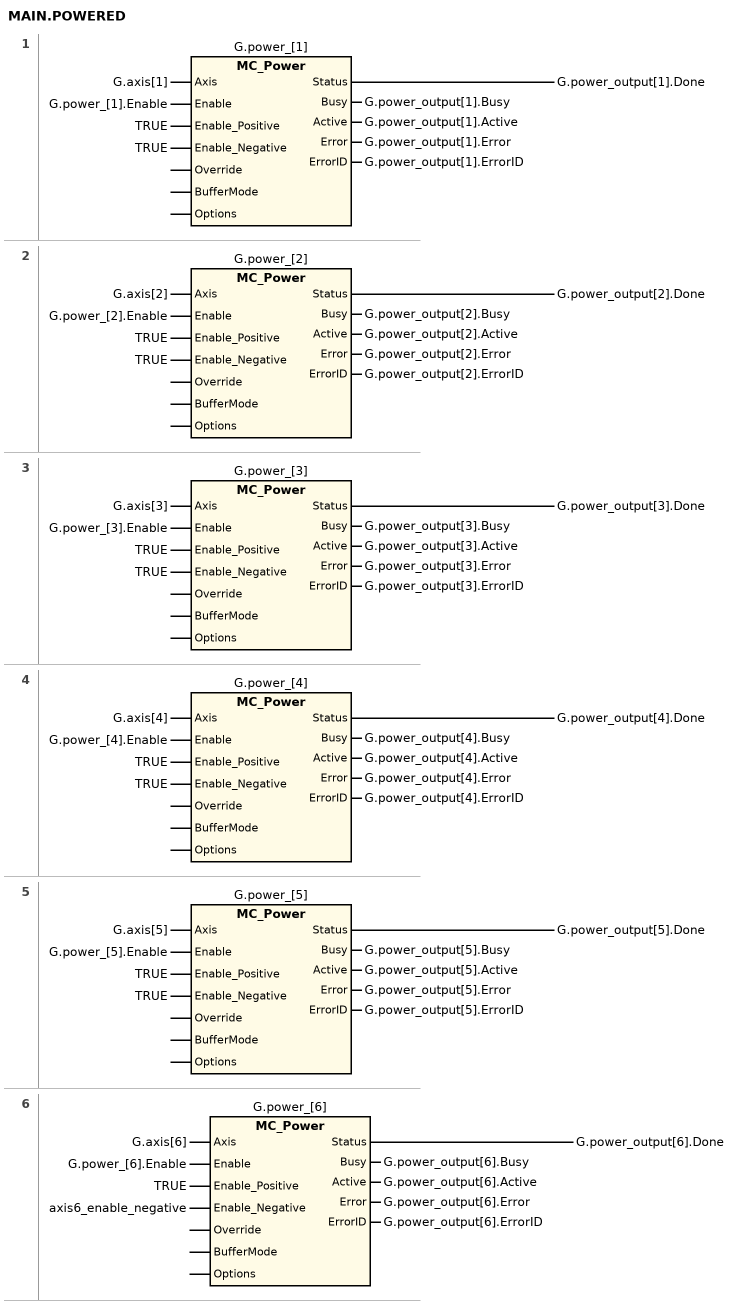
// NETWORK 1
G.power_[1](
    Axis := G.axis[1],
    Enable := G.power_[1].Enable,
    Enable_Positive := TRUE,
    Enable_Negative := TRUE,
    Busy => G.power_output[1].Busy,
    Active => G.power_output[1].Active,
    Error => G.power_output[1].Error,
    ErrorID => G.power_output[1].ErrorID); // MC_Power
G.power_output[1].Done := G.power_[1].Status;

// NETWORK 2
G.power_[2](
    Axis := G.axis[2],
    Enable := G.power_[2].Enable,
    Enable_Positive := TRUE,
    Enable_Negative := TRUE,
    Busy => G.power_output[2].Busy,
    Active => G.power_output[2].Active,
    Error => G.power_output[2].Error,
    ErrorID => G.power_output[2].ErrorID); // MC_Power
G.power_output[2].Done := G.power_[2].Status;

// NETWORK 3
G.power_[3](
    Axis := G.axis[3],
    Enable := G.power_[3].Enable,
    Enable_Positive := TRUE,
    Enable_Negative := TRUE,
    Busy => G.power_output[3].Busy,
    Active => G.power_output[3].Active,
    Error => G.power_output[3].Error,
    ErrorID => G.power_output[3].ErrorID); // MC_Power
G.power_output[3].Done := G.power_[3].Status;

// NETWORK 4
G.power_[4](
    Axis := G.axis[4],
    Enable := G.power_[4].Enable,
    Enable_Positive := TRUE,
    Enable_Negative := TRUE,
    Busy => G.power_output[4].Busy,
    Active => G.power_output[4].Active,
    Error => G.power_output[4].Error,
    ErrorID => G.power_output[4].ErrorID); // MC_Power
G.power_output[4].Done := G.power_[4].Status;

// NETWORK 5
G.power_[5](
    Axis := G.axis[5],
    Enable := G.power_[5].Enable,
    Enable_Positive := TRUE,
    Enable_Negative := TRUE,
    Busy => G.power_output[5].Busy,
    Active => G.power_output[5].Active,
    Error => G.power_output[5].Error,
    ErrorID => G.power_output[5].ErrorID); // MC_Power
G.power_output[5].Done := G.power_[5].Status;

// NETWORK 6
G.power_[6](
    Axis := G.axis[6],
    Enable := G.power_[6].Enable,
    Enable_Positive := TRUE,
    Enable_Negative := axis6_enable_negative,
    Busy => G.power_output[6].Busy,
    Active => G.power_output[6].Active,
    Error => G.power_output[6].Error,
    ErrorID => G.power_output[6].ErrorID); // MC_Power
G.power_output[6].Done := G.power_[6].Status;

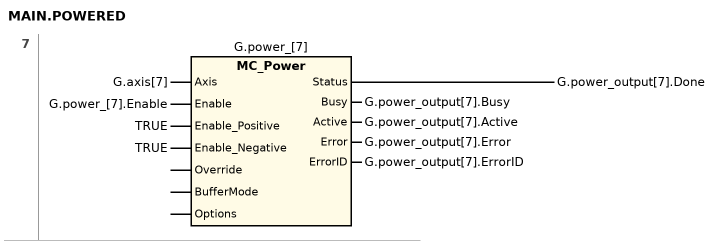
// NETWORK 7
G.power_[7](
    Axis := G.axis[7],
    Enable := G.power_[7].Enable,
    Enable_Positive := TRUE,
    Enable_Negative := TRUE,
    Busy => G.power_output[7].Busy,
    Active => G.power_output[7].Active,
    Error => G.power_output[7].Error,
    ErrorID => G.power_output[7].ErrorID); // MC_Power
G.power_output[7].Done := G.power_[7].Status;
END_ACTION

ACTION RESETED:
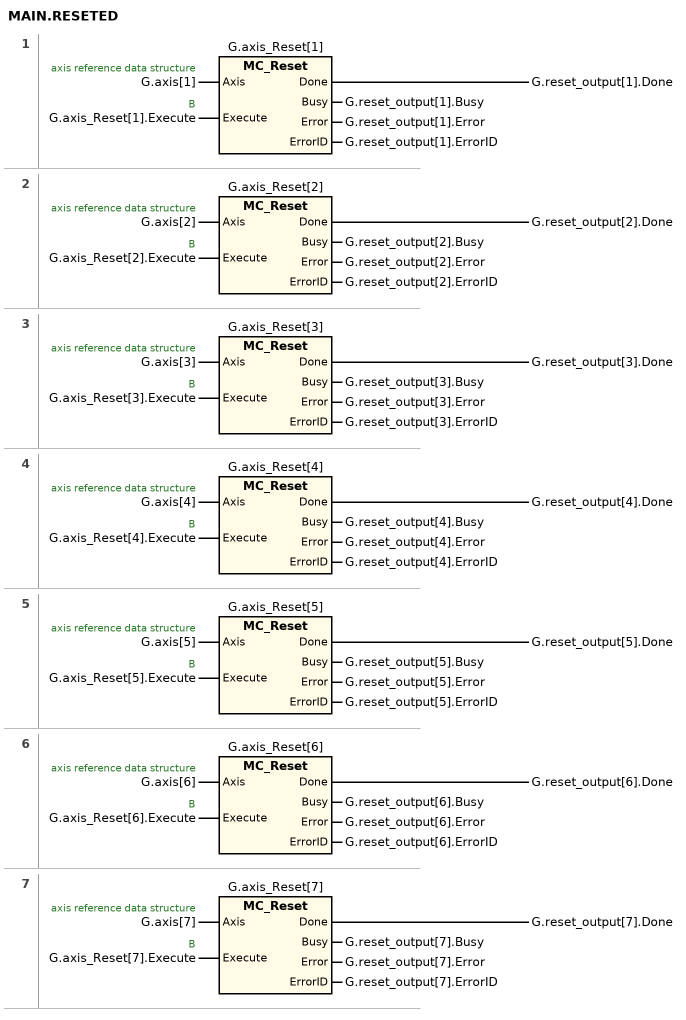
// NETWORK 1
//   G.axis[1]: axis reference data structure
//   G.axis_Reset[1].Execute: B
G.axis_Reset[1](
    Axis := G.axis[1],
    Execute := G.axis_Reset[1].Execute,
    Busy => G.reset_output[1].Busy,
    Error => G.reset_output[1].Error,
    ErrorID => G.reset_output[1].ErrorID); // MC_Reset
G.reset_output[1].Done := G.axis_Reset[1].Done;

// NETWORK 2
//   G.axis[2]: axis reference data structure
//   G.axis_Reset[2].Execute: B
G.axis_Reset[2](
    Axis := G.axis[2],
    Execute := G.axis_Reset[2].Execute,
    Busy => G.reset_output[2].Busy,
    Error => G.reset_output[2].Error,
    ErrorID => G.reset_output[2].ErrorID); // MC_Reset
G.reset_output[2].Done := G.axis_Reset[2].Done;

// NETWORK 3
//   G.axis[3]: axis reference data structure
//   G.axis_Reset[3].Execute: B
G.axis_Reset[3](
    Axis := G.axis[3],
    Execute := G.axis_Reset[3].Execute,
    Busy => G.reset_output[3].Busy,
    Error => G.reset_output[3].Error,
    ErrorID => G.reset_output[3].ErrorID); // MC_Reset
G.reset_output[3].Done := G.axis_Reset[3].Done;

// NETWORK 4
//   G.axis[4]: axis reference data structure
//   G.axis_Reset[4].Execute: B
G.axis_Reset[4](
    Axis := G.axis[4],
    Execute := G.axis_Reset[4].Execute,
    Busy => G.reset_output[4].Busy,
    Error => G.reset_output[4].Error,
    ErrorID => G.reset_output[4].ErrorID); // MC_Reset
G.reset_output[4].Done := G.axis_Reset[4].Done;

// NETWORK 5
//   G.axis[5]: axis reference data structure
//   G.axis_Reset[5].Execute: B
G.axis_Reset[5](
    Axis := G.axis[5],
    Execute := G.axis_Reset[5].Execute,
    Busy => G.reset_output[5].Busy,
    Error => G.reset_output[5].Error,
    ErrorID => G.reset_output[5].ErrorID); // MC_Reset
G.reset_output[5].Done := G.axis_Reset[5].Done;

// NETWORK 6
//   G.axis[6]: axis reference data structure
//   G.axis_Reset[6].Execute: B
G.axis_Reset[6](
    Axis := G.axis[6],
    Execute := G.axis_Reset[6].Execute,
    Busy => G.reset_output[6].Busy,
    Error => G.reset_output[6].Error,
    ErrorID => G.reset_output[6].ErrorID); // MC_Reset
G.reset_output[6].Done := G.axis_Reset[6].Done;

// NETWORK 7
//   G.axis[7]: axis reference data structure
//   G.axis_Reset[7].Execute: B
G.axis_Reset[7](
    Axis := G.axis[7],
    Execute := G.axis_Reset[7].Execute,
    Busy => G.reset_output[7].Busy,
    Error => G.reset_output[7].Error,
    ErrorID => G.reset_output[7].ErrorID); // MC_Reset
G.reset_output[7].Done := G.axis_Reset[7].Done;
END_ACTION

ACTION SETPOSITIONGEN:
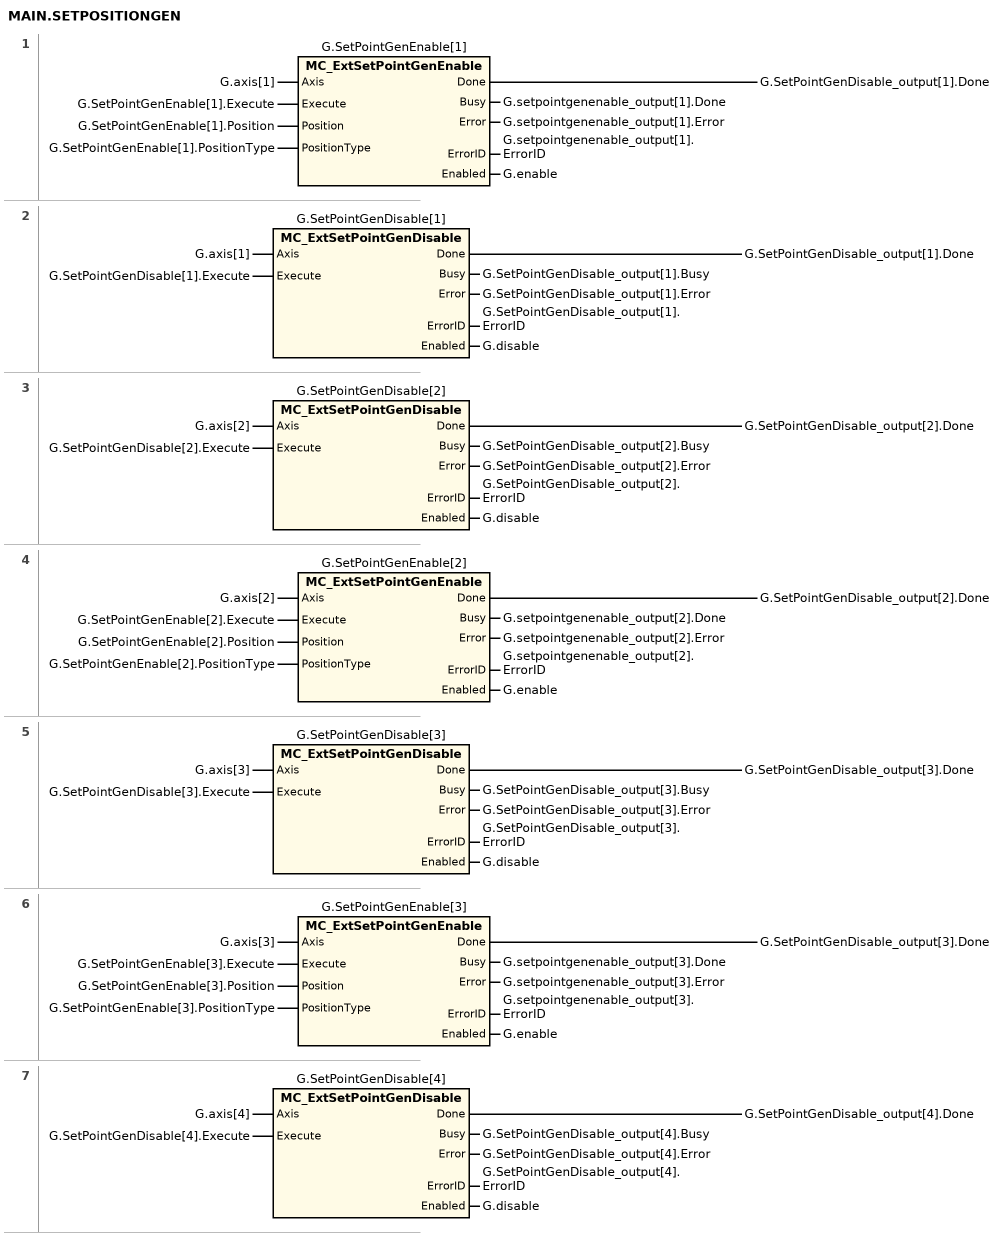
// NETWORK 1
G.SetPointGenEnable[1](
    Axis := G.axis[1],
    Execute := G.SetPointGenEnable[1].Execute,
    Position := G.SetPointGenEnable[1].Position,
    PositionType := G.SetPointGenEnable[1].PositionType,
    Busy => G.setpointgenenable_output[1].Done,
    Error => G.setpointgenenable_output[1].Error,
    ErrorID => G.setpointgenenable_output[1].ErrorID,
    Enabled => G.enable); // MC_ExtSetPointGenEnable
G.SetPointGenDisable_output[1].Done := G.SetPointGenEnable[1].Done;

// NETWORK 2
G.SetPointGenDisable[1](
    Axis := G.axis[1],
    Execute := G.SetPointGenDisable[1].Execute,
    Busy => G.SetPointGenDisable_output[1].Busy,
    Error => G.SetPointGenDisable_output[1].Error,
    ErrorID => G.SetPointGenDisable_output[1].ErrorID,
    Enabled => G.disable); // MC_ExtSetPointGenDisable
G.SetPointGenDisable_output[1].Done := G.SetPointGenDisable[1].Done;

// NETWORK 3
G.SetPointGenDisable[2](
    Axis := G.axis[2],
    Execute := G.SetPointGenDisable[2].Execute,
    Busy => G.SetPointGenDisable_output[2].Busy,
    Error => G.SetPointGenDisable_output[2].Error,
    ErrorID => G.SetPointGenDisable_output[2].ErrorID,
    Enabled => G.disable); // MC_ExtSetPointGenDisable
G.SetPointGenDisable_output[2].Done := G.SetPointGenDisable[2].Done;

// NETWORK 4
G.SetPointGenEnable[2](
    Axis := G.axis[2],
    Execute := G.SetPointGenEnable[2].Execute,
    Position := G.SetPointGenEnable[2].Position,
    PositionType := G.SetPointGenEnable[2].PositionType,
    Busy => G.setpointgenenable_output[2].Done,
    Error => G.setpointgenenable_output[2].Error,
    ErrorID => G.setpointgenenable_output[2].ErrorID,
    Enabled => G.enable); // MC_ExtSetPointGenEnable
G.SetPointGenDisable_output[2].Done := G.SetPointGenEnable[2].Done;

// NETWORK 5
G.SetPointGenDisable[3](
    Axis := G.axis[3],
    Execute := G.SetPointGenDisable[3].Execute,
    Busy => G.SetPointGenDisable_output[3].Busy,
    Error => G.SetPointGenDisable_output[3].Error,
    ErrorID => G.SetPointGenDisable_output[3].ErrorID,
    Enabled => G.disable); // MC_ExtSetPointGenDisable
G.SetPointGenDisable_output[3].Done := G.SetPointGenDisable[3].Done;

// NETWORK 6
G.SetPointGenEnable[3](
    Axis := G.axis[3],
    Execute := G.SetPointGenEnable[3].Execute,
    Position := G.SetPointGenEnable[3].Position,
    PositionType := G.SetPointGenEnable[3].PositionType,
    Busy => G.setpointgenenable_output[3].Done,
    Error => G.setpointgenenable_output[3].Error,
    ErrorID => G.setpointgenenable_output[3].ErrorID,
    Enabled => G.enable); // MC_ExtSetPointGenEnable
G.SetPointGenDisable_output[3].Done := G.SetPointGenEnable[3].Done;

// NETWORK 7
G.SetPointGenDisable[4](
    Axis := G.axis[4],
    Execute := G.SetPointGenDisable[4].Execute,
    Busy => G.SetPointGenDisable_output[4].Busy,
    Error => G.SetPointGenDisable_output[4].Error,
    ErrorID => G.SetPointGenDisable_output[4].ErrorID,
    Enabled => G.disable); // MC_ExtSetPointGenDisable
G.SetPointGenDisable_output[4].Done := G.SetPointGenDisable[4].Done;

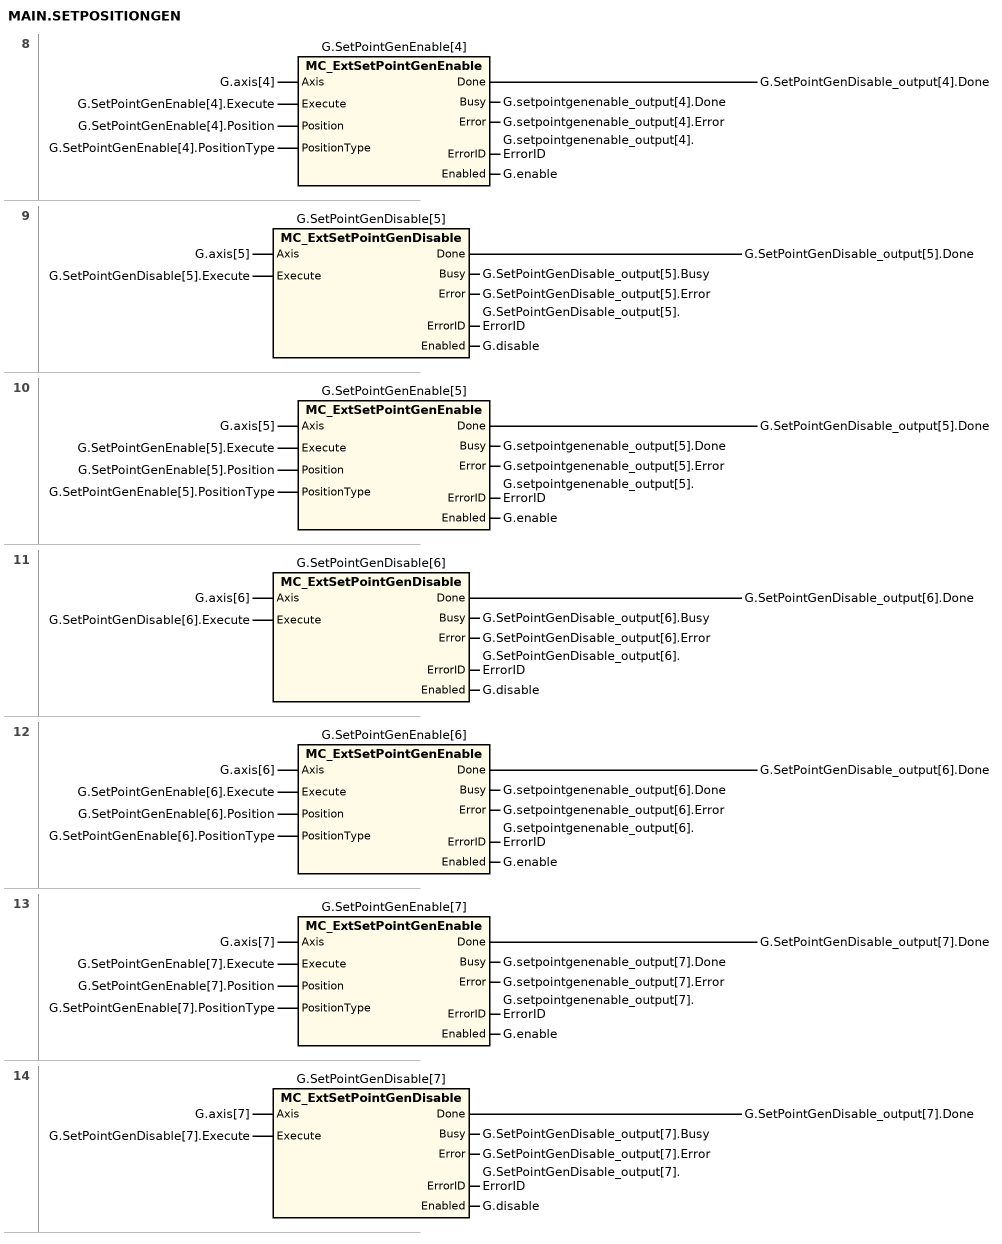
// NETWORK 8
G.SetPointGenEnable[4](
    Axis := G.axis[4],
    Execute := G.SetPointGenEnable[4].Execute,
    Position := G.SetPointGenEnable[4].Position,
    PositionType := G.SetPointGenEnable[4].PositionType,
    Busy => G.setpointgenenable_output[4].Done,
    Error => G.setpointgenenable_output[4].Error,
    ErrorID => G.setpointgenenable_output[4].ErrorID,
    Enabled => G.enable); // MC_ExtSetPointGenEnable
G.SetPointGenDisable_output[4].Done := G.SetPointGenEnable[4].Done;

// NETWORK 9
G.SetPointGenDisable[5](
    Axis := G.axis[5],
    Execute := G.SetPointGenDisable[5].Execute,
    Busy => G.SetPointGenDisable_output[5].Busy,
    Error => G.SetPointGenDisable_output[5].Error,
    ErrorID => G.SetPointGenDisable_output[5].ErrorID,
    Enabled => G.disable); // MC_ExtSetPointGenDisable
G.SetPointGenDisable_output[5].Done := G.SetPointGenDisable[5].Done;

// NETWORK 10
G.SetPointGenEnable[5](
    Axis := G.axis[5],
    Execute := G.SetPointGenEnable[5].Execute,
    Position := G.SetPointGenEnable[5].Position,
    PositionType := G.SetPointGenEnable[5].PositionType,
    Busy => G.setpointgenenable_output[5].Done,
    Error => G.setpointgenenable_output[5].Error,
    ErrorID => G.setpointgenenable_output[5].ErrorID,
    Enabled => G.enable); // MC_ExtSetPointGenEnable
G.SetPointGenDisable_output[5].Done := G.SetPointGenEnable[5].Done;

// NETWORK 11
G.SetPointGenDisable[6](
    Axis := G.axis[6],
    Execute := G.SetPointGenDisable[6].Execute,
    Busy => G.SetPointGenDisable_output[6].Busy,
    Error => G.SetPointGenDisable_output[6].Error,
    ErrorID => G.SetPointGenDisable_output[6].ErrorID,
    Enabled => G.disable); // MC_ExtSetPointGenDisable
G.SetPointGenDisable_output[6].Done := G.SetPointGenDisable[6].Done;

// NETWORK 12
G.SetPointGenEnable[6](
    Axis := G.axis[6],
    Execute := G.SetPointGenEnable[6].Execute,
    Position := G.SetPointGenEnable[6].Position,
    PositionType := G.SetPointGenEnable[6].PositionType,
    Busy => G.setpointgenenable_output[6].Done,
    Error => G.setpointgenenable_output[6].Error,
    ErrorID => G.setpointgenenable_output[6].ErrorID,
    Enabled => G.enable); // MC_ExtSetPointGenEnable
G.SetPointGenDisable_output[6].Done := G.SetPointGenEnable[6].Done;

// NETWORK 13
G.SetPointGenEnable[7](
    Axis := G.axis[7],
    Execute := G.SetPointGenEnable[7].Execute,
    Position := G.SetPointGenEnable[7].Position,
    PositionType := G.SetPointGenEnable[7].PositionType,
    Busy => G.setpointgenenable_output[7].Done,
    Error => G.setpointgenenable_output[7].Error,
    ErrorID => G.setpointgenenable_output[7].ErrorID,
    Enabled => G.enable); // MC_ExtSetPointGenEnable
G.SetPointGenDisable_output[7].Done := G.SetPointGenEnable[7].Done;

// NETWORK 14
G.SetPointGenDisable[7](
    Axis := G.axis[7],
    Execute := G.SetPointGenDisable[7].Execute,
    Busy => G.SetPointGenDisable_output[7].Busy,
    Error => G.SetPointGenDisable_output[7].Error,
    ErrorID => G.SetPointGenDisable_output[7].ErrorID,
    Enabled => G.disable); // MC_ExtSetPointGenDisable
G.SetPointGenDisable_output[7].Done := G.SetPointGenDisable[7].Done;
END_ACTION

END_PROGRAM

// ---- POUs/init.TcPOU
FUNCTION_BLOCK init
VAR_INPUT
END_VAR
VAR_OUTPUT
END_VAR
VAR
	i:INT;
	step:INT:=0;
	init_watchdog : TON;
	all_powered : BOOL;
END_VAR

(*
FUNCTION_BLOCK: init
功能说明:
  上电初始化流程：给 7 轴上电(MC_Power)，等待 Done；若超时或出现错误则进入 _err。

状态机(step):
  0) 进入初始化：清理控制命令，启动看门狗
  1) 等待上电完成：检测 Done/错误/超时并跳转
*)

CASE step OF
0:
	// 进入 init 的第一个周期：清理边沿触发量，避免上一次状态遗留导致重复触发
	FOR i:=1 TO 7 DO
		G.SetPointGenEnable[i].Execute := FALSE;
		G.SetPointGenDisable[i].Execute := FALSE;
		G.axis_Reset[i].Execute := FALSE;
		G.power_[i].Enable := TRUE;
	END_FOR
	G.self_check_done := FALSE;
	G.startup_loading_ready := FALSE;
	G.selfcheck_reset_req := TRUE;

	init_watchdog(IN:=TRUE, PT:=T#5S);
	step := 1;

1:
	// 持续保持上电请求，并监控上电结果
	FOR i:=1 TO 7 DO
		G.power_[i].Enable := TRUE;

		// 若任一轴出现错误：进入 _err(安全态)，避免 init/reset 来回震荡
		IF G.axis[i].Status.Error OR G.power_output[i].Error THEN
			init_watchdog(IN:=FALSE);
			step := 0;
			G.gen_state := _err;
			RETURN;
		END_IF
	END_FOR

	// 等待上电全部完成
	all_powered := TRUE;
	FOR i:=1 TO 7 DO
		IF NOT G.power_output[i].Done THEN
			all_powered := FALSE;
		END_IF
	END_FOR

	// 超时保护：上电迟迟不完成，进入 _err(安全态)
	init_watchdog(IN:=TRUE);
	IF init_watchdog.Q THEN
		init_watchdog(IN:=FALSE);
		step := 0;
		G.gen_state := _err;
		RETURN;
	END_IF

	// 上电全部完成：记录各轴当前绝对位置作为 init_pos(用于绝对->相对转换)，进入自检
	IF all_powered THEN
		FOR i:=1 TO 7 DO
			G.init_pos[i] := G.axis[i].NcToPlc.ActPos;
		END_FOR
		init_watchdog(IN:=FALSE);
		step := 0;
		G.gen_state := _self_check;
	END_IF
END_CASE

END_FUNCTION_BLOCK

// ---- POUs/handle.TcPOU
FUNCTION_BLOCK handle
VAR_INPUT
END_VAR
VAR_OUTPUT
END_VAR
VAR
	i,j,k:INT;
    handoff : Handoff;
    handoff_reinit : BOOL;
	v_step		: LREAL;
	avg_window	: INT;
	avg_window_size : INT := 20;
	return_handoff_bypass : BOOL;

	act_hh		:	ARRAY[1..7] OF ARRAY [1..30] OF LREAL;
	pos_abs		:	LREAL;
	legacy_vel	:	LREAL;

	init_wait : TON;
	init_retry : ARRAY[1..7] OF UINT;
	init_drop : ARRAY[1..7] OF BOOL;
	return_wait : ARRAY[1..7] OF TON;
	return_wait_state : ARRAY[1..7] OF INT;
	return_enable_retry : ARRAY[1..7] OF UINT;
	return_enable_drop : ARRAY[1..7] OF BOOL;
	return_clear_stop : ARRAY[1..7] OF MC_Stop;
	return_clear_stop_active : ARRAY[1..7] OF BOOL;
	axis4_wait : TON;
	axis4_wait_state : INT;
	axis4_retry : UINT;
	axis4_drop : BOOL;
	init_done : BOOL := FALSE;
	all_enabled : BOOL;
	all_powered : BOOL;
	has_axis_error : BOOL;
	hold_active : BOOL := FALSE;

	// 上位机通信看门狗。超时锁存后只能通过显式恢复握手解除。
	host_watchdog_timer : TON;
	host_last_session_id : UDINT := 0;
	host_last_heartbeat_sequence : UDINT := 0;
	host_heartbeat_seen : BOOL := FALSE;
	host_session_changed : BOOL;
	host_heartbeat_changed : BOOL;
	host_timeout_latched : BOOL := FALSE;
	host_timeout_prev : BOOL := FALSE;
	// 看门狗超时后锁存一次外部设定值保持位置。
	// 不能每拍把 Actual Position 回写为下一拍设定值，否则编码器微动会被回灌到 NC。
	host_hold_abs : ARRAY[1..7] OF LREAL;
	host_hold_captured : BOOL := FALSE;
	host_all_stopped : BOOL;
	host_return_stop_active : ARRAY[1..7] OF BOOL;
	host_return_stop_exec : ARRAY[1..7] OF BOOL;
	host_axis4_stop_active : BOOL := FALSE;
	fb_host_return_stop : ARRAY[1..7] OF MC_Stop;

	right_slimit : ARRAY[1..7] OF LREAL;
	slimit_enable : ARRAY[1..7] OF BOOL := [TRUE, FALSE, TRUE, FALSE, TRUE, TRUE, FALSE];

	ext_setpoint_enabled : ARRAY[1..7] OF BOOL := [FALSE,FALSE,FALSE,FALSE,FALSE,FALSE,FALSE];
	spg_enable_exec	: ARRAY[1..7] OF BOOL;
	spg_disable_exec : ARRAY[1..7] OF BOOL;

	return_enable : ARRAY[1..7] OF BOOL := [TRUE, FALSE, FALSE, FALSE, FALSE, TRUE, FALSE];
	return_state : ARRAY[1..7] OF INT;
	return_exec : ARRAY[1..7] OF BOOL;
	return_target_abs : ARRAY[1..7] OF LREAL;
	return_velocity : ARRAY[1..7] OF LREAL;
	return_acc : ARRAY[1..7] OF LREAL;
	return_dec : ARRAY[1..7] OF LREAL;
	return_jerk : ARRAY[1..7] OF LREAL;
	return_finish_error : ARRAY[1..7] OF BOOL;
	return_error_id_pending : ARRAY[1..7] OF UDINT;
	fb_return_move_abs : ARRAY[1..7] OF MC_MoveAbsolute;

	axis4_manual_state : INT := 0;
	axis4_request_dir_now : INT := 0;
	axis4_requested_dir : INT := 0;
	axis4_pending_dir : INT := 0;
	axis4_move_exec : BOOL := FALSE;
	axis4_stop_exec : BOOL := FALSE;
	axis4_finish_error : BOOL := FALSE;
	axis4_error_id_pending : UDINT := 0;
	axis4_manual_velocity : LREAL := 60;
	axis4_manual_acc : LREAL := 200;
	axis4_manual_dec : LREAL := 200;
	axis4_manual_jerk : LREAL := 500.0;
	axis4_manual_direction : MC_Direction := MC_Direction.MC_Positive_Direction;
	fb_axis4_move_velocity : MC_MoveVelocity;
	fb_axis4_stop : MC_Stop;
	ramp_counter: ARRAY[1..7] OF INT;
	act_h_prev : ARRAY[1..7] OF LREAL;

	traj_pos     : ARRAY[1..7] OF LREAL;
	traj_vel     : ARRAY[1..7] OF LREAL;
	traj_acc     : ARRAY[1..7] OF LREAL;
	acc_raw      : LREAL;

	traj_wn      : LREAL := 60.0;
	traj_vmax    : ARRAY[1..7] OF LREAL := [80, 0, 80, 0, 80, 80, 0];
	traj_amax    : ARRAY[1..7] OF LREAL := [2000, 0, 2000, 0, 2000, 2000, 0];
	traj_enable  : ARRAY[1..7] OF BOOL := [TRUE, FALSE, TRUE, FALSE, TRUE, TRUE, FALSE];
END_VAR

host_session_changed := G.host_session_id <> host_last_session_id;
host_heartbeat_changed := host_session_changed OR
	(G.host_heartbeat_sequence <> host_last_heartbeat_sequence);

IF host_session_changed THEN
	// 非零会话发生变化表示新的上位机接管，必须重新完成恢复握手。
	IF host_last_session_id <> 0 THEN
		host_timeout_latched := TRUE;
	END_IF
	host_last_session_id := G.host_session_id;
END_IF

IF host_heartbeat_changed THEN
	host_last_heartbeat_sequence := G.host_heartbeat_sequence;
END_IF

host_heartbeat_seen := G.host_session_id <> 0;
// 心跳变化的扫描周期将 TON 复位；序号连续 2s 不变化才判定通信超时。
host_watchdog_timer(
	IN:=host_heartbeat_seen AND NOT host_heartbeat_changed,
	PT:=T#2S
);
IF (NOT host_heartbeat_seen) OR host_watchdog_timer.Q THEN
	host_timeout_latched := TRUE;
END_IF
IF G.host_comm_timeout THEN
	host_timeout_latched := TRUE;
END_IF
G.host_comm_timeout := host_timeout_latched;

handoff_reinit := G.handle_reinit_req;
IF G.handle_reinit_req THEN
	init_done := FALSE;
	init_wait(IN:=FALSE);
	axis4_wait(IN:=FALSE);
	axis4_retry := 0;
	axis4_drop := FALSE;
	G.handle_reinit_done := FALSE;
	G.handle_reinit_req := FALSE;

	FOR i:=1 TO 7 DO
		ext_setpoint_enabled[i] := FALSE;
		spg_enable_exec[i] := FALSE;
		spg_disable_exec[i] := FALSE;
		init_retry[i] := 0;
		init_drop[i] := FALSE;
		return_wait[i](IN:=FALSE);
		return_enable_retry[i] := 0;
		return_enable_drop[i] := FALSE;
		return_clear_stop_active[i] := FALSE;
		return_state[i] := 0;
		return_exec[i] := FALSE;
		return_finish_error[i] := FALSE;
		return_error_id_pending[i] := 0;
		traj_pos[i] := 0.0;
		traj_vel[i] := 0.0;
		traj_acc[i] := 0.0;
		host_hold_abs[i] := 0.0;
		handoff.leg_cmd[i].Req := FALSE;
		handoff.leg_cmd[i].Busy := FALSE;
		handoff.leg_cmd[i].Done := FALSE;
		handoff.leg_cmd[i].Error := FALSE;
		handoff.leg_cmd[i].ErrorId := 0;
	END_FOR
	host_hold_captured := FALSE;
	host_timeout_prev := FALSE;

	axis4_manual_state := 0;
	axis4_request_dir_now := 0;
	axis4_requested_dir := 0;
	axis4_pending_dir := 0;
	axis4_move_exec := FALSE;
	axis4_stop_exec := FALSE;
	axis4_finish_error := FALSE;
	axis4_error_id_pending := 0;
	G.axis4_fwd_req := FALSE;
	G.axis4_rev_req := FALSE;
	G.axis4_manual_busy := FALSE;
	G.axis4_manual_done := FALSE;
	G.axis4_manual_error := FALSE;
	G.axis4_manual_error_id := 0;
END_IF

all_powered := TRUE;
FOR i:=1 TO 7 DO
	IF NOT G.power_output[i].Done THEN
		all_powered := FALSE;
		EXIT;
	END_IF
END_FOR

has_axis_error := FALSE;
FOR i:=1 TO 7 DO
	IF G.axis[i].Status.Error OR G.power_output[i].Error OR G.reset_output[i].Error THEN
		has_axis_error := TRUE;
		EXIT;
	END_IF
END_FOR

handoff(ready:=init_done AND all_powered AND NOT has_axis_error AND NOT G.host_comm_timeout AND NOT handoff_reinit,
    interrupted:=NOT all_powered OR has_axis_error OR G.host_comm_timeout OR handoff_reinit);

IF (NOT all_powered) OR has_axis_error THEN
	// 在自动清错、重建参考和重启 Power 之前保留故障当拍，恢复后不清除。
	G.estop_diag_host_timeout := G.host_comm_timeout;
	FOR j:=1 TO 7 DO
		G.estop_diag_axis[j] := G.axis[j].Status;
		G.estop_diag_power[j] := G.power_output[j];
		G.estop_diag_reset[j] := G.reset_output[j];
		G.estop_diag_power_enable[j] := G.power_[j].Enable;
		G.estop_diag_power_positive[j] := G.power_[j].Enable_Positive;
		G.estop_diag_power_negative[j] := G.power_[j].Enable_Negative;
		G.estop_diag_return_state[j] := return_state[j];
		G.estop_diag_return_cmd[j] := handoff.leg_cmd[j];
		G.estop_diag_move_error[j] := fb_return_move_abs[j].Error;
		G.estop_diag_move_aborted[j] := fb_return_move_abs[j].CommandAborted;
		G.estop_diag_move_error_id[j] := fb_return_move_abs[j].ErrorID;
		G.estop_diag_enable_error[j] := G.SetPointGenEnable[j].Error;
		G.estop_diag_enable_error_id[j] := G.SetPointGenEnable[j].ErrorID;
		G.estop_diag_disable_error[j] := G.SetPointGenDisable[j].Error;
		G.estop_diag_disable_error_id[j] := G.SetPointGenDisable[j].ErrorID;
		G.estop_diag_act_pos[j] := G.axis[j].NcToPlc.ActPos;
		G.estop_diag_act_vel[j] := G.axis[j].NcToPlc.ActVelo;
		G.estop_diag_feed_pos[j] := G.axis[j].PlcToNc.ExtSetPos;
		G.estop_diag_feed_vel[j] := G.axis[j].PlcToNc.ExtSetVelo;
		G.estop_diag_refer_abs[j] := G.refer[j] + G.init_pos[j];
	END_FOR
	G.estop_diag_count := G.estop_diag_count + 1;
	G.estop_hold_req := TRUE;
	FOR j:=1 TO 7 DO
		G.SetPointGenDisable[j].Execute := FALSE;
		G.Act_pos[j] := G.axis[j].NcToPlc.ActPos - G.init_pos[j];
		G.act_pos_from_left[j] := G.axis[j].NcToPlc.ActPos - G.leftlimit[j];
		G.refer[j] := G.Act_pos[j];
		G.ref_slow[j] := G.Act_pos[j];
		G.act_h[j] := G.Act_pos[j];
		G.act_hf[j] := G.Act_pos[j];
		G.refer_from_left[j] := G.act_pos_from_left[j];
		FOR k:=1 TO 30 DO
			act_hh[j][k] := G.Act_pos[j];
		END_FOR
		act_h_prev[j] := G.Act_pos[j];
		traj_pos[j] := G.Act_pos[j];
		traj_vel[j] := 0.0;
		traj_acc[j] := 0.0;
	END_FOR

	G.gen_state := _err;
	RETURN;
END_IF

IF NOT init_done THEN
	init_wait(IN:=TRUE, PT:=G.recovery_wait_timeout);
	IF init_wait.Q THEN
		G.gen_state := _err;
		G.estop_hold_req := TRUE;
		init_wait(IN:=FALSE);
		RETURN;
	END_IF
	all_enabled := TRUE;
	FOR i:=1 TO 7 DO
		G.SetPointGenEnable[i].Execute := TRUE;
		IF init_drop[i] THEN
			init_drop[i] := FALSE;
		ELSIF G.SetPointGenEnable[i].Error THEN
			IF init_retry[i] < G.recovery_max_retries THEN
				G.SetPointGenEnable[i].Execute := FALSE;
				init_drop[i] := TRUE;
				init_retry[i] := init_retry[i] + 1;
			END_IF
		END_IF
		IF NOT G.SetPointGenEnable[i].Done OR G.SetPointGenEnable[i].Error THEN
			all_enabled := FALSE;
		END_IF
	END_FOR

	IF all_enabled THEN
		FOR j:=1 TO 7 DO
			G.Act_pos[j] := G.axis[j].NcToPlc.ActPos - G.init_pos[j];
			G.act_pos_from_left[j] := G.axis[j].NcToPlc.ActPos - G.leftlimit[j];
			G.ref_slow[j] := G.Act_pos[j];
			G.act_h[j] := G.Act_pos[j];
			G.act_hf[j] := G.Act_pos[j];
			G.refer[j] := G.Act_pos[j];
			G.refer_from_left[j] := G.act_pos_from_left[j];
			ext_setpoint_enabled[j] := TRUE;

			FOR k:=1 TO 30 DO
				act_hh[j][k] := G.Act_pos[j];
			END_FOR
			act_h_prev[j] := G.Act_pos[j];
			traj_pos[j] := G.Act_pos[j];
			traj_vel[j] := 0.0;
			traj_acc[j] := 0.0;
			IF slimit_enable[j] THEN
				right_slimit[j] := G.leftlimit[j] + G.rslimit_distance[j];
			END_IF
			handoff.leg_cmd[j].Busy := FALSE;
			handoff.leg_cmd[j].Done := FALSE;
			handoff.leg_cmd[j].Error := FALSE;
			handoff.leg_cmd[j].ErrorId := 0;
		END_FOR

		G.axis4_manual_busy := FALSE;
		G.axis4_manual_done := FALSE;
		G.axis4_manual_error := FALSE;
		G.axis4_manual_error_id := 0;

		init_wait(IN:=FALSE);
		init_done := TRUE;
		// 通信超时未解除时不提前确认恢复；正式握手后会再次进入本初始化流程。
		G.handle_reinit_done := NOT G.host_comm_timeout;
	END_IF
	RETURN;
END_IF


IF G.host_comm_timeout THEN
	G.handle_reinit_done := FALSE;

	IF (NOT host_timeout_prev) OR (NOT host_hold_captured) THEN
		// 仅在进入超时保持时采样一次。之后始终维持同一绝对位置，
		// 避免 Actual -> Set Position 的逐周期回灌导致低频来回摆动。
		FOR i:=1 TO 7 DO
			host_hold_abs[i] := G.axis[i].NcToPlc.ActPos;
		END_FOR
		host_hold_captured := TRUE;
	END_IF

	IF NOT host_timeout_prev THEN
		// 仅捕获超时发生时已经在运行的独立运动，禁止恢复后自动续跑。
		FOR i:=1 TO 7 DO
			host_return_stop_active[i] := return_enable[i] AND
				((return_state[i] <> 0) OR handoff.leg_cmd[i].Busy OR fb_return_move_abs[i].Busy);
			host_return_stop_exec[i] := FALSE;
		END_FOR
		host_axis4_stop_active := (axis4_manual_state <> 0) OR fb_axis4_move_velocity.Busy;
	END_IF

	// 超时期间持续清除运动请求，避免上位机重连时把旧请求重新送入状态机。


	G.axis4_fwd_req := FALSE;
	G.axis4_rev_req := FALSE;

	axis4_move_exec := FALSE;
	host_all_stopped := TRUE;

	FOR i:=1 TO 7 DO
		spg_enable_exec[i] := FALSE;
		spg_disable_exec[i] := FALSE;
		return_exec[i] := FALSE;
		handoff.leg_cmd[i].Req := FALSE;
		handoff.leg_cmd[i].Done := FALSE;

		// 实际位置仍实时刷新用于诊断；外部参考始终保持超时边沿的锁存位置。
		G.Act_pos[i] := G.axis[i].NcToPlc.ActPos - G.init_pos[i];
		G.act_pos_from_left[i] := G.axis[i].NcToPlc.ActPos - G.leftlimit[i];
		G.refer[i] := host_hold_abs[i] - G.init_pos[i];
		G.ref_slow[i] := G.refer[i];
		G.act_h[i] := G.refer[i];
		G.act_hf[i] := G.refer[i];
		G.refer_from_left[i] := host_hold_abs[i] - G.leftlimit[i];
		FOR k:=1 TO 30 DO
			act_hh[i][k] := G.refer[i];
		END_FOR
		act_h_prev[i] := G.refer[i];
		traj_pos[i] := G.refer[i];
		traj_vel[i] := 0.0;
		traj_acc[i] := 0.0;

		IF host_return_stop_active[i] THEN
			IF fb_host_return_stop[i].Done THEN
				host_return_stop_exec[i] := FALSE;
				host_return_stop_active[i] := FALSE;
			ELSIF fb_host_return_stop[i].Error THEN
				// 拉低一个扫描周期清除错误，下一周期继续尝试受控停止。
				host_return_stop_exec[i] := FALSE;
				host_all_stopped := FALSE;
			ELSE
				host_return_stop_exec[i] := TRUE;
				host_all_stopped := FALSE;
			END_IF
		ELSE
			host_return_stop_exec[i] := FALSE;
		END_IF
		handoff.leg_cmd[i].Busy := host_return_stop_active[i];

		IF ext_setpoint_enabled[i] THEN
			MC_ExtSetPointGenFeed(
				Position:=host_hold_abs[i],
				Velocity:=0.0,
				Acceleration:=0.0,
				Direction:=1,
				Axis:=G.axis[i]);
		END_IF

		// 所有运动功能块在看门狗分支中仍保持每扫描调用。
		G.SetPointGenEnable[i].Execute := FALSE;
		G.SetPointGenDisable[i].Execute := FALSE;
		fb_return_move_abs[i](
			Axis:=G.axis[i],
			Position:=return_target_abs[i],
			Velocity:=return_velocity[i],
			Acceleration:=return_acc[i],
			Deceleration:=return_dec[i],
			Jerk:=return_jerk[i],
			Execute:=FALSE
		);
		fb_host_return_stop[i](
			Axis:=G.axis[i],
			Execute:=host_return_stop_exec[i],
			Deceleration:=4000.0,
			Jerk:=10000.0
		);
	END_FOR

	IF host_axis4_stop_active THEN
		IF fb_axis4_stop.Done THEN
			axis4_stop_exec := FALSE;
			host_axis4_stop_active := FALSE;
		ELSIF fb_axis4_stop.Error THEN
			// 拉低一个扫描周期清除错误，下一周期继续尝试受控停止。
			axis4_stop_exec := FALSE;
			host_all_stopped := FALSE;
		ELSE
			axis4_stop_exec := TRUE;
			host_all_stopped := FALSE;
		END_IF
	ELSE
		axis4_stop_exec := FALSE;
	END_IF
	G.axis4_manual_busy := host_axis4_stop_active;
	G.axis4_manual_done := FALSE;

	fb_axis4_move_velocity(
		Axis:=G.axis[4],
		Execute:=FALSE,
		Velocity:=axis4_manual_velocity,
		Acceleration:=axis4_manual_acc,
		Deceleration:=axis4_manual_dec,
		Jerk:=axis4_manual_jerk,
		Direction:=axis4_manual_direction
	);
	fb_axis4_stop(
		Axis:=G.axis[4],
		Execute:=axis4_stop_exec,
		Deceleration:=axis4_manual_dec,
		Jerk:=axis4_manual_jerk
	);

	// 清请求并解除超时即为 PLC 对恢复请求的确认；随后复用既有重初始化流程。
	IF G.host_recover_req AND host_heartbeat_seen AND
		(NOT host_watchdog_timer.Q) AND host_all_stopped THEN
		host_timeout_latched := FALSE;
		G.host_comm_timeout := FALSE;
		G.host_recover_req := FALSE;
		G.handle_reinit_req := TRUE;
	END_IF

	host_timeout_prev := G.host_comm_timeout;
	RETURN;
END_IF

host_timeout_prev := FALSE;
host_hold_captured := FALSE;
// 非超时状态收到的恢复请求没有业务含义，清除以免成为下一次超时的陈旧握手。
G.host_recover_req := FALSE;

G.estop_hold_req := FALSE;

IF G.cylinder5_press_req THEN
	G.cylinder5_value := 500;
ELSE
	G.cylinder5_value := 2000;
END_IF

FOR i:=1 TO 7 DO
	spg_enable_exec[i] := FALSE;
	spg_disable_exec[i] := FALSE;
	return_exec[i] := FALSE;
END_FOR
axis4_move_exec := FALSE;
axis4_stop_exec := FALSE;

FOR j:=1 TO 7 DO
	G.Act_pos[j] := G.axis[j].NcToPlc.ActPos - G.init_pos[j];
	G.act_pos_from_left[j] := G.axis[j].NcToPlc.ActPos - G.leftlimit[j];
	G.refer_from_left[j] := (G.refer[j] + G.init_pos[j]) - G.leftlimit[j];

	// 事务运动开始后直到接管，参与轴的参考由PLC独占。
	// 状态 30/31 期间冻结参考输入，防止驱动层接收矛盾信号（禁用→重启 同时 参考变化）
	IF return_enable[j] AND handoff.freeze[j] THEN
		G.refer[j] := traj_pos[j];
		G.refer_from_left[j] := traj_pos[j] + G.init_pos[j] - G.leftlimit[j];
		CONTINUE;
	END_IF

	v_step := G.v_limit[j];
	// 回退接管旁路：回退 Busy 期间跳过斜坡/均值，避免回退末端重新进入慢链路
	return_handoff_bypass := handoff.freeze[j];
	IF return_handoff_bypass THEN
		avg_window := 1;
		ramp_counter[j] := 0;
	ELSE
		ramp_counter[j] := MIN(ramp_counter[j] + 1, avg_window_size);
		avg_window := MAX(1, ramp_counter[j]);
	END_IF

	FOR k:=2 TO 20 DO
		act_hh[j][22-k] := act_hh[j][21-k];
	END_FOR

	IF slimit_enable[j] THEN
		IF (G.axis[j].NcToPlc.ActPos >= right_slimit[j]) AND (G.refer[j] > G.ref_slow[j]) THEN
			G.refer[j] := G.ref_slow[j];
		END_IF
	END_IF

	IF return_handoff_bypass THEN
		G.ref_slow[j] := G.refer[j];
	ELSIF (G.refer[j] - G.ref_slow[j]) > v_step THEN
		G.ref_slow[j] := G.ref_slow[j] + v_step;
	ELSIF (G.refer[j] - G.ref_slow[j]) < -v_step THEN
		G.ref_slow[j] := G.ref_slow[j] - v_step;
	ELSE
		G.ref_slow[j] := G.refer[j];
	END_IF

	IF return_handoff_bypass THEN
		FOR i:=1 TO 20 DO
			act_hh[j][i] := G.ref_slow[j];
		END_FOR
		G.act_h[j] := G.ref_slow[j];
	ELSE
		act_hh[j][1] := G.ref_slow[j];
		G.act_h[j] := 0;
		FOR i:=1 TO avg_window DO
			G.act_h[j] := G.act_h[j] + act_hh[j][i] / TO_LREAL(avg_window);
		END_FOR
	END_IF

	IF traj_enable[j] AND NOT return_handoff_bypass THEN
		acc_raw := traj_wn * traj_wn * (G.refer[j] - traj_pos[j]) - 2.0 * traj_wn * traj_vel[j];
		IF acc_raw > traj_amax[j] THEN
			acc_raw := traj_amax[j];
		ELSIF acc_raw < -traj_amax[j] THEN
			acc_raw := -traj_amax[j];
		END_IF
		traj_acc[j] := acc_raw;
		traj_vel[j] := traj_vel[j] + 0.001 * traj_acc[j];
		IF traj_vel[j] > traj_vmax[j] THEN
			traj_vel[j] := traj_vmax[j];
		ELSIF traj_vel[j] < -traj_vmax[j] THEN
			traj_vel[j] := -traj_vmax[j];
		END_IF
		traj_pos[j] := traj_pos[j] + 0.001 * traj_vel[j];
		IF ABS(G.refer[j] - traj_pos[j]) < 0.001 AND ABS(traj_vel[j]) < 0.01 THEN
			traj_pos[j] := G.refer[j];
			traj_vel[j] := 0.0;
			traj_acc[j] := 0.0;
		END_IF
	ELSE
		traj_pos[j] := G.act_h[j];
		traj_vel[j] := 0.0;
		traj_acc[j] := 0.0;
	END_IF
END_FOR

FOR i:=1 TO 7 DO
	IF NOT return_enable[i] THEN
		CONTINUE;
	END_IF

	IF return_state[i] = 0 THEN
		handoff.leg_cmd[i].Busy := FALSE;
		IF NOT handoff.leg_cmd[i].Req THEN
			handoff.leg_cmd[i].Done := FALSE;
			handoff.leg_cmd[i].Error := FALSE;
			handoff.leg_cmd[i].ErrorId := 0;
			return_finish_error[i] := FALSE;
			return_error_id_pending[i] := 0;
		ELSIF (NOT handoff.leg_cmd[i].Done) AND (NOT handoff.leg_cmd[i].Error) THEN
			// 子流程请求由Handoff发起；运动参数仅在此锁存一次。
			return_target_abs[i] := handoff.leg_cmd[i].TargetAbs;
			return_velocity[i] := handoff.leg_cmd[i].Velocity;
			return_acc[i] := handoff.leg_cmd[i].Acc;
			return_dec[i] := handoff.leg_cmd[i].Dec;
			return_jerk[i] := handoff.leg_cmd[i].Jerk;
			return_state[i] := 10;
		END_IF
	END_IF

    IF return_wait_state[i] <> return_state[i] THEN
        return_wait[i](IN:=FALSE);
        return_wait_state[i] := return_state[i];
    END_IF
    return_wait[i](IN:=(return_state[i] = 10) OR (return_state[i] = 20) OR (return_state[i] = 31), PT:=G.recovery_wait_timeout);
	IF return_state[i] <> 31 THEN
		return_enable_retry[i] := 0;
		return_enable_drop[i] := FALSE;
	END_IF
	IF ((return_state[i] = 10) OR (return_state[i] = 20)) AND
		(handoff.abort_motion OR G.SetPointGenDisable[i].Error OR return_wait[i].Q) THEN
		return_clear_stop_active[i] := return_state[i] = 20;
		return_finish_error[i] := TRUE;
        handoff.leg_error[i] := G.handoff_err_timeout;
        IF G.SetPointGenDisable[i].Error THEN handoff.leg_error[i] := G.handoff_err_disable; END_IF
        IF handoff.abort_motion THEN handoff.leg_error[i] := G.handoff_err_move; END_IF
        return_error_id_pending[i] := G.SetPointGenDisable[i].ErrorID;
        handoff.leg_cmd[i].Error := TRUE;
        handoff.leg_cmd[i].ErrorId := return_error_id_pending[i];
		return_state[i] := 30;
	END_IF
	CASE return_state[i] OF
	10:
		handoff.leg_cmd[i].Busy := TRUE;
		spg_disable_exec[i] := TRUE;
		IF G.SetPointGenDisable[i].Done OR NOT G.SetPointGenDisable[i].Enabled THEN
			ext_setpoint_enabled[i] := FALSE;
			return_state[i] := 20;
		END_IF

	20:
		handoff.leg_cmd[i].Busy := TRUE;
		return_exec[i] := TRUE;
		G.refer_from_left[i] := return_target_abs[i] - G.leftlimit[i];

		// 接近目标不能代替功能块完成确认，否则未启动或被中断的命令也会被当成成功。
		IF handoff.abort_motion OR fb_return_move_abs[i].Error OR fb_return_move_abs[i].CommandAborted THEN
			return_finish_error[i] := TRUE;
			return_error_id_pending[i] := fb_return_move_abs[i].ErrorID;
            return_clear_stop_active[i] := TRUE;
            handoff.leg_error[i] := G.handoff_err_move;
            handoff.leg_cmd[i].Error := TRUE;
            handoff.leg_cmd[i].ErrorId := return_error_id_pending[i];
			return_state[i] := 30;
		ELSIF fb_return_move_abs[i].Done THEN
			return_finish_error[i] := FALSE;
			return_error_id_pending[i] := 0;
			return_state[i] := 30;
		END_IF

	30:
		handoff.leg_cmd[i].Busy := TRUE;
		IF (ABS(G.axis[i].NcToPlc.ActVelo) <= 0.5) AND NOT return_clear_stop_active[i] THEN
			G.Act_pos[i] := G.axis[i].NcToPlc.ActPos - G.init_pos[i];
			G.act_pos_from_left[i] := G.axis[i].NcToPlc.ActPos - G.leftlimit[i];
            // 停稳后只对齐一次；下一扫描先预送，再重新使能。
            G.refer[i] := G.Act_pos[i];
            G.ref_slow[i] := G.Act_pos[i];
            G.act_h[i] := G.Act_pos[i];
            G.act_hf[i] := G.Act_pos[i];
            G.refer_from_left[i] := G.act_pos_from_left[i];
            FOR k:=1 TO 30 DO act_hh[i][k] := G.Act_pos[i]; END_FOR
            act_h_prev[i] := G.Act_pos[i];
            traj_pos[i] := G.Act_pos[i];
			traj_vel[i] := 0.0;
			traj_acc[i] := 0.0;
			// 先留出一个完整 PLC 扫描周期预送当前设定值，再重新使能外部设定值发生器。
			return_state[i] := 31;
		END_IF

	31:
		handoff.leg_cmd[i].Busy := TRUE;
		spg_enable_exec[i] := TRUE;
		IF return_wait[i].Q THEN
			G.gen_state := _err;
			G.estop_hold_req := TRUE;
			RETURN;
		END_IF
		IF return_enable_drop[i] THEN
			return_enable_drop[i] := FALSE;
		ELSIF G.SetPointGenEnable[i].Error THEN
			IF return_enable_retry[i] < G.recovery_max_retries THEN
				spg_enable_exec[i] := FALSE;
				return_enable_drop[i] := TRUE;
				return_enable_retry[i] := return_enable_retry[i] + 1;
			END_IF
		END_IF
		IF G.SetPointGenEnable[i].Done AND NOT G.SetPointGenEnable[i].Error THEN
			ext_setpoint_enabled[i] := TRUE;
			handoff.leg_cmd[i].Busy := FALSE;
			IF return_finish_error[i] THEN
				handoff.leg_cmd[i].Done := FALSE;
				handoff.leg_cmd[i].Error := TRUE;
				handoff.leg_cmd[i].ErrorId := return_error_id_pending[i];
			ELSE
				handoff.leg_cmd[i].Done := TRUE;
				handoff.leg_cmd[i].Error := FALSE;
				handoff.leg_cmd[i].ErrorId := 0;
			END_IF
			return_finish_error[i] := FALSE;
			return_error_id_pending[i] := 0;
			return_state[i] := 0;
		END_IF
	END_CASE
END_FOR

axis4_request_dir_now := 0;
IF G.axis4_fwd_req AND NOT G.axis4_rev_req THEN
	axis4_request_dir_now := 1;
ELSIF G.axis4_rev_req AND NOT G.axis4_fwd_req THEN
	axis4_request_dir_now := -1;
END_IF

IF axis4_manual_state = 0 THEN
	G.axis4_manual_busy := FALSE;
	IF axis4_request_dir_now = 0 THEN
		G.axis4_manual_done := FALSE;
		G.axis4_manual_error := FALSE;
		G.axis4_manual_error_id := 0;
	ELSIF NOT G.axis4_manual_error THEN
		G.axis4_manual_done := FALSE;
		G.axis4_manual_error := FALSE;
		G.axis4_manual_error_id := 0;
		axis4_requested_dir := axis4_request_dir_now;
		axis4_pending_dir := 0;
		axis4_finish_error := FALSE;
		axis4_error_id_pending := 0;
		axis4_manual_state := 10;
	END_IF
END_IF

IF axis4_wait_state <> axis4_manual_state THEN
	axis4_wait(IN:=FALSE);
	axis4_wait_state := axis4_manual_state;
	axis4_retry := 0;
	axis4_drop := FALSE;
END_IF
axis4_wait(IN:=(axis4_manual_state = 10) OR (axis4_manual_state = 30) OR (axis4_manual_state = 40), PT:=G.recovery_wait_timeout);
IF axis4_wait.Q THEN
	IF axis4_manual_state = 40 THEN
		G.gen_state := _err;
		G.estop_hold_req := TRUE;
		RETURN;
	ELSE
		axis4_finish_error := TRUE;
		axis4_error_id_pending := G.SetPointGenDisable[4].ErrorID;
		axis4_pending_dir := 0;
		axis4_manual_state := 40;
		axis4_wait(IN:=FALSE);
	END_IF
END_IF
CASE axis4_manual_state OF
10:
	G.axis4_manual_busy := TRUE;
	spg_disable_exec[4] := TRUE;
	IF axis4_drop THEN
		axis4_drop := FALSE;
	ELSIF G.SetPointGenDisable[4].Error THEN
		IF axis4_retry < G.recovery_max_retries THEN
			spg_disable_exec[4] := FALSE;
			axis4_drop := TRUE;
			axis4_retry := axis4_retry + 1;
		ELSE
			axis4_finish_error := TRUE;
			axis4_error_id_pending := G.SetPointGenDisable[4].ErrorID;
			axis4_manual_state := 40;
		END_IF
	END_IF
	IF NOT G.SetPointGenDisable[4].Error AND (G.SetPointGenDisable[4].Done OR NOT G.SetPointGenDisable[4].Enabled) THEN
		ext_setpoint_enabled[4] := FALSE;
		axis4_manual_state := 20;
	END_IF

20:
	G.axis4_manual_busy := TRUE;
	axis4_pending_dir := axis4_request_dir_now;
	IF axis4_requested_dir >= 0 THEN
		axis4_manual_direction := MC_Direction.MC_Positive_Direction;
	ELSE
		axis4_manual_direction := MC_Direction.MC_Negative_Direction;
	END_IF

	IF axis4_pending_dir = 0 THEN
		axis4_manual_state := 30;
	ELSIF axis4_pending_dir <> axis4_requested_dir THEN
		axis4_manual_state := 30;
	ELSE
		axis4_move_exec := TRUE;
	END_IF

	IF fb_axis4_move_velocity.Error THEN
		axis4_finish_error := TRUE;
		axis4_error_id_pending := fb_axis4_move_velocity.ErrorID;
		G.axis4_manual_error_id := fb_axis4_move_velocity.ErrorID;
		axis4_pending_dir := 0;
		axis4_manual_state := 40;
	ELSIF fb_axis4_move_velocity.CommandAborted THEN
		// 被 MC_Stop 中止属于正常方向切换，进入停稳流程，不锁存为错误。
		axis4_pending_dir := axis4_request_dir_now;
		axis4_manual_state := 30;
	END_IF

30:
	G.axis4_manual_busy := TRUE;
	axis4_pending_dir := axis4_request_dir_now;
	axis4_stop_exec := TRUE;

    IF axis4_drop THEN
        axis4_drop := FALSE;
    ELSIF fb_axis4_stop.Error THEN
        IF axis4_retry < G.recovery_max_retries THEN
            axis4_stop_exec := FALSE;
            axis4_drop := TRUE;
            axis4_retry := axis4_retry + 1;
        ELSE
            axis4_finish_error := TRUE;
            axis4_error_id_pending := fb_axis4_stop.ErrorID;
            axis4_pending_dir := 0;
            axis4_manual_state := 40;
        END_IF
    END_IF
    IF NOT fb_axis4_stop.Error AND (fb_axis4_stop.Done OR (ABS(G.axis[4].NcToPlc.ActVelo) <= 0.05)) THEN
		// 无论是否还有请求，先经过状态39释放 MC_Stop 一个完整扫描周期。
		axis4_manual_state := 39;
	END_IF

39:
	G.axis4_manual_busy := TRUE;
	// MC_Stop 需要一个 Execute=FALSE 的完整周期，
	// 再重新触发 MoveVelocity 或 SetPointGenEnable。
	axis4_pending_dir := axis4_request_dir_now;
	IF (axis4_pending_dir <> 0) AND NOT axis4_finish_error THEN
		axis4_requested_dir := axis4_pending_dir;
		axis4_manual_state := 20;
	ELSE
		axis4_requested_dir := 0;
		axis4_manual_state := 40;
	END_IF

40:
	G.axis4_manual_busy := TRUE;
	G.Act_pos[4] := G.axis[4].NcToPlc.ActPos - G.init_pos[4];
	G.act_pos_from_left[4] := G.axis[4].NcToPlc.ActPos - G.leftlimit[4];
	G.refer[4] := G.Act_pos[4];
	G.ref_slow[4] := G.Act_pos[4];
	G.act_h[4] := G.Act_pos[4];
	G.act_hf[4] := G.Act_pos[4];
	G.refer_from_left[4] := G.act_pos_from_left[4];
	FOR k:=1 TO 30 DO
		act_hh[4][k] := G.Act_pos[4];
	END_FOR
	act_h_prev[4] := G.Act_pos[4];
	traj_pos[4] := G.Act_pos[4];
	traj_vel[4] := 0.0;
	traj_acc[4] := 0.0;
	spg_enable_exec[4] := TRUE;
	IF axis4_drop THEN
		axis4_drop := FALSE;
	ELSIF G.SetPointGenEnable[4].Error THEN
		IF axis4_retry < G.recovery_max_retries THEN
			spg_enable_exec[4] := FALSE;
			axis4_drop := TRUE;
			axis4_retry := axis4_retry + 1;
		ELSE
			G.gen_state := _err;
			G.estop_hold_req := TRUE;
			RETURN;
		END_IF
	END_IF
	IF G.SetPointGenEnable[4].Done AND NOT G.SetPointGenEnable[4].Error THEN
		ext_setpoint_enabled[4] := TRUE;
		G.axis4_manual_busy := FALSE;
		IF axis4_finish_error THEN
			G.axis4_manual_done := FALSE;
			G.axis4_manual_error := TRUE;
			G.axis4_manual_error_id := axis4_error_id_pending;
		ELSE
			G.axis4_manual_done := TRUE;
			G.axis4_manual_error := FALSE;
			G.axis4_manual_error_id := 0;
		END_IF
		axis4_finish_error := FALSE;
		axis4_error_id_pending := 0;
		axis4_manual_state := 0;
	END_IF
END_CASE

FOR i:=1 TO 7 DO
	IF G.power_output[i].Error THEN
		G.axis_Reset[i].Execute := TRUE;
	END_IF
END_FOR

FOR i:=1 TO 7 DO
	// 计划回退结束后，状态 31 的预送周期和 SetPointGenEnable 过渡周期都必须喂入当前设定值。
	// 否则 NC 重新接管时会短暂使用禁用前遗留的左窗口设定值，造成约一个窗口宽度的反向尖峰。
	IF ext_setpoint_enabled[i] OR (return_state[i] = 31) OR spg_enable_exec[i] THEN
		IF traj_enable[i] THEN
			pos_abs := traj_pos[i] + G.init_pos[i];
			MC_ExtSetPointGenFeed(
				Position     := pos_abs,
				Velocity     := traj_vel[i],
				Acceleration := traj_acc[i],
				Direction    := 1,
				Axis         := G.axis[i]);
		ELSE
			pos_abs := G.act_h[i] + G.init_pos[i];
			legacy_vel := (G.act_h[i] - act_h_prev[i]) / 0.001;
			MC_ExtSetPointGenFeed(
				Position     := pos_abs,
				Velocity     := legacy_vel,
				Acceleration := 0,
				Direction    := 1,
				Axis         := G.axis[i]);
		END_IF
		G.act_hf[i] := G.act_h[i];
	ELSE
		G.act_hf[i] := G.axis[i].NcToPlc.ActPos - G.init_pos[i];
	END_IF
	act_h_prev[i] := G.act_h[i];
END_FOR

FOR i:=1 TO 7 DO
	G.SetPointGenEnable[i].Execute := spg_enable_exec[i];
	G.SetPointGenDisable[i].Execute := spg_disable_exec[i];
	return_clear_stop[i](Axis:=G.axis[i], Execute:=return_clear_stop_active[i],
		Deceleration:=return_dec[i], Jerk:=return_jerk[i]);
	IF return_clear_stop_active[i] AND return_clear_stop[i].Done THEN
		return_clear_stop_active[i] := FALSE;
	END_IF
	fb_return_move_abs[i](
		Axis:=G.axis[i],
		Position:=return_target_abs[i],
		Velocity:=return_velocity[i],
		Acceleration:=return_acc[i],
		Deceleration:=return_dec[i],
		Jerk:=return_jerk[i],
		Execute:=return_exec[i]
	);
END_FOR

fb_axis4_move_velocity(
	Axis:=G.axis[4],
	Execute:=axis4_move_exec,
	Velocity:=axis4_manual_velocity,
	Acceleration:=axis4_manual_acc,
	Deceleration:=axis4_manual_dec,
	Jerk:=axis4_manual_jerk,
	Direction:=axis4_manual_direction
);
fb_axis4_stop(
	Axis:=G.axis[4],
	Execute:=axis4_stop_exec,
	Deceleration:=axis4_manual_dec,
	Jerk:=axis4_manual_jerk
);

END_FUNCTION_BLOCK

// ---- POUs/Handoff.TcPOU
FUNCTION_BLOCK Handoff
VAR_INPUT
    ready : BOOL;
    interrupted : BOOL;
    // handle内部子流程回写状态；不向ADS上位机公开触发接口。
    leg_cmd : ARRAY[1..7] OF ST_AxisPlannedReturnCmd;
    leg_error : ARRAY[1..7] OF UDINT;
END_VAR
VAR_OUTPUT
    freeze : ARRAY[1..7] OF BOOL;
    abort_motion : BOOL;
END_VAR
VAR
    latched : ST_HandoffCmd;
    active_id : UDINT;
    last_request : UDINT;
    active : BOOL;
    interrupted_pending : BOOL;
    initialized : BOOL;
    was_ready : BOOL;
    fault_code : UDINT;
    fault_axis : INT;
    fault_nc : UDINT;
    outputs : ARRAY[1..4] OF WORD;
    tick : UDINT;
    phase_start : UDINT;
    motion_start : UDINT;
    motion_recorded : ARRAY[1..2] OF BOOL;
    phase : INT;
    previous_phase : INT;
    next_phase : INT;
    wait_slot : INT;
    wait_max : UDINT;
    elapsed : UDINT;
    slot, axis_index, holder, mover, i : INT;
    participates, all_finished, params_valid : BOOL;
END_VAR

// 本功能块每个1ms任务扫描调用一次；不依赖ADS快照或上位机周期。
tick := tick + 1;
previous_phase := phase;
next_phase := phase;
IF NOT initialized THEN
    outputs[1] := G.cylinder1_value;
    outputs[2] := G.cylinder2_value;
    outputs[3] := G.cylinder3_value;
    outputs[4] := G.cylinder4_value;
    IF ready THEN
        G.cyl_cmd := outputs;
        initialized := TRUE;
    END_IF
END_IF

IF ready AND NOT was_ready AND NOT active THEN
    G.cyl_cmd[1] := G.cylinder1_value;
    G.cyl_cmd[2] := G.cylinder2_value;
    G.cyl_cmd[3] := G.cylinder3_value;
    G.cyl_cmd[4] := G.cylinder4_value;
END_IF
was_ready := ready;

IF active AND interrupted THEN
    interrupted_pending := TRUE;
    fault_code := G.handoff_err_interrupted;
    fault_axis := 0;
    fault_nc := 0;
    abort_motion := TRUE;
END_IF

IF (G.handoff_cmd.request_id <> 0) AND (G.handoff_cmd.request_id <> G.handoff_status.ack_id) AND (G.handoff_cmd.request_id <> last_request) AND NOT (active AND (G.handoff_cmd.request_id = active_id)) THEN
    last_request := G.handoff_cmd.request_id;
    params_valid := (G.handoff_cmd.leg_mask = 1) OR (G.handoff_cmd.leg_mask = 2) OR (G.handoff_cmd.leg_mask = 3);
    FOR slot := 1 TO 2 DO
        participates := (G.handoff_cmd.leg_mask = 3) OR (G.handoff_cmd.leg_mask = slot);
        IF participates THEN
            params_valid := params_valid AND (G.handoff_cmd.velocity[slot] > 0) AND (G.handoff_cmd.acc[slot] > 0);
        END_IF
    END_FOR
    IF active OR NOT ready OR NOT params_valid OR (((G.handoff_cmd.leg_mask AND 1) <> 0) AND leg_cmd[1].Busy) OR (((G.handoff_cmd.leg_mask AND 2) <> 0) AND leg_cmd[6].Busy) THEN
        G.handoff_status.ack_id := last_request;
        G.handoff_status.done_id := last_request;
        G.handoff_status.result := 2;
        G.handoff_status.error_code := G.handoff_err_rejected;
        G.handoff_status.error_axis := 0;
        IF active THEN G.handoff_status.reject_reason := 1;
        ELSIF NOT ready THEN G.handoff_status.reject_reason := 2;
        ELSE G.handoff_status.reject_reason := 3; END_IF
    ELSE
        latched := G.handoff_cmd;
        active_id := latched.request_id;
        active := TRUE;
        abort_motion := FALSE;
        interrupted_pending := FALSE;
        fault_code := 0;
        fault_axis := 0;
        fault_nc := 0;
        G.handoff_status.ack_id := active_id;
        G.handoff_status.done_id := 0;
        G.handoff_status.result := 0;
        G.handoff_status.error_code := 0;
        G.handoff_status.error_axis := 0;
        G.handoff_status.nc_error_code := 0;
        G.handoff_status.reject_reason := 0;
        G.handoff_status.leg_mask := latched.leg_mask;
        FOR i := 1 TO 8 DO G.handoff_status.phase_ms[i] := 0; END_FOR
        FOR i := 1 TO 7 DO
            leg_cmd[i].Req := FALSE;
            leg_error[i] := 0;
        END_FOR
        FOR slot := 1 TO 2 DO motion_recorded[slot] := FALSE; END_FOR
        outputs[1] := G.cyl_cmd[1];
        outputs[2] := G.cyl_cmd[2];
        outputs[3] := G.cyl_cmd[3];
        outputs[4] := G.cyl_cmd[4];
        next_phase := 10;
    END_IF
END_IF

IF active AND ready AND NOT interrupted THEN
    IF interrupted_pending THEN
        // 原停轴/重初始化路径已完成；恢复后只执行夹爪收尾，不续跑旧目标。
        interrupted_pending := FALSE;
        next_phase := 40;
        FOR i := 1 TO 7 DO leg_cmd[i].Req := FALSE; END_FOR
    ELSE
        elapsed := tick - phase_start;
        CASE phase OF
        10, 20, 40, 50:
            wait_slot := 1;
            IF phase = 20 THEN wait_slot := 2; END_IF
            IF phase = 40 THEN wait_slot := 3; END_IF
            IF phase = 50 THEN wait_slot := 4; END_IF
            wait_max := 0;
            FOR slot := 1 TO 2 DO
                IF (latched.leg_mask = 3) OR (latched.leg_mask = slot) THEN
                    wait_max := MAX(wait_max, latched.wait_ms[slot][wait_slot]);
                END_IF
            END_FOR
            IF elapsed >= wait_max THEN next_phase := phase + 10; END_IF
        30:
            all_finished := TRUE;
            FOR slot := 1 TO 2 DO
                IF (latched.leg_mask = 3) OR (latched.leg_mask = slot) THEN
                    axis_index := 1;
                    IF slot = 2 THEN axis_index := 6; END_IF
                    IF leg_error[axis_index] <> 0 THEN
                        abort_motion := TRUE;
                        IF fault_code = 0 THEN
                            fault_code := leg_error[axis_index];
                            fault_axis := axis_index;
                            fault_nc := leg_cmd[axis_index].ErrorId;
                        END_IF
                    END_IF
                    IF leg_cmd[axis_index].Busy OR NOT (leg_cmd[axis_index].Done OR leg_cmd[axis_index].Error) THEN
                        all_finished := FALSE;
                    ELSIF NOT motion_recorded[slot] THEN
                        G.handoff_status.phase_ms[5 + slot] := tick - motion_start;
                        motion_recorded[slot] := TRUE;
                    END_IF
                END_IF
            END_FOR
            IF all_finished THEN next_phase := 40; END_IF
        60:
            IF G.handoff_takeover_id = active_id THEN
                // 移交时写回当前输出，屏蔽事务期间残留的上位机电缸命令。
                G.cyl_cmd := outputs;
                next_phase := 0;
                active := FALSE;
                abort_motion := FALSE;
            END_IF
        END_CASE
    END_IF
END_IF

IF next_phase <> phase THEN
    IF phase = 10 THEN G.handoff_status.phase_ms[1] := tick - phase_start; END_IF
    IF phase = 20 THEN G.handoff_status.phase_ms[2] := tick - phase_start; END_IF
    IF phase = 30 THEN G.handoff_status.phase_ms[3] := tick - phase_start; END_IF
    IF phase = 40 THEN G.handoff_status.phase_ms[4] := tick - phase_start; END_IF
    IF phase = 50 THEN G.handoff_status.phase_ms[5] := tick - phase_start; END_IF
    phase := next_phase;
    phase_start := tick;
    G.handoff_status.phase := phase;
    G.handoff_status.phase_seq := G.handoff_status.phase_seq + 1;
    IF phase = 30 THEN motion_start := tick; END_IF
    IF phase = 60 THEN
        G.handoff_status.ack_id := active_id;
        G.handoff_status.done_id := active_id;
        G.handoff_status.error_code := fault_code;
        G.handoff_status.error_axis := fault_axis;
        G.handoff_status.nc_error_code := fault_nc;
        G.handoff_status.reject_reason := 0;
        IF fault_code = 0 THEN G.handoff_status.result := 1;
        ELSE G.handoff_status.result := 2; END_IF
    END_IF
END_IF

FOR slot := 1 TO 2 DO
    axis_index := 1;
    IF slot = 2 THEN axis_index := 6; END_IF
    participates := active AND ((latched.leg_mask = 3) OR (latched.leg_mask = slot));
    freeze[axis_index] := participates AND (phase >= 30);
    IF participates AND ready AND NOT interrupted AND NOT interrupted_pending THEN
        holder := slot * 2 - 1;
        mover := slot * 2;
        IF (phase = 10) OR (phase = 40) THEN
            outputs[holder] := latched.cyl_clamp[holder];
            outputs[mover] := latched.cyl_clamp[mover];
        ELSIF (phase = 20) OR (phase = 30) THEN
            outputs[holder] := latched.cyl_clamp[holder];
            outputs[mover] := latched.cyl_open[mover];
        ELSIF phase = 50 THEN
            outputs[holder] := latched.cyl_open[holder];
            outputs[mover] := latched.cyl_clamp[mover];
        END_IF
        leg_cmd[axis_index].Req := phase = 30;
        IF (phase = 30) AND (previous_phase <> 30) THEN
            leg_cmd[axis_index].TargetAbs := latched.target_abs[slot];
            leg_cmd[axis_index].Velocity := latched.velocity[slot];
            leg_cmd[axis_index].Acc := latched.acc[slot];
            leg_cmd[axis_index].Dec := latched.dec[slot];
            leg_cmd[axis_index].Jerk := latched.jerk[slot];
        END_IF
    END_IF
END_FOR
IF NOT active AND ready THEN outputs := G.cyl_cmd; END_IF
// 非_handle时自检等原有流程仍直接控制电缸，事务保留内部输出直到恢复。
IF G.gen_state = _handle THEN
    G.cylinder1_value := outputs[1];
    G.cylinder2_value := outputs[2];
    G.cylinder3_value := outputs[3];
    G.cylinder4_value := outputs[4];
END_IF

END_FUNCTION_BLOCK

// ---- POUs/clear_err.TcPOU
FUNCTION_BLOCK clear_err
VAR_INPUT
END_VAR
VAR_OUTPUT
END_VAR
VAR
	i:INT;
	step:INT:=0;
	settle_timer:TON;
	all_powered:BOOL;
	has_err:BOOL;
END_VAR

(* 
Post-error recovery:
  - keep the handle input frozen
  - cold start or a fresh _init cycle must return to _init until self-check is completed
  - otherwise wait until errors are gone and all axes are powered again
  - then reinitialize handle references from the current position
*)

has_err := FALSE;
FOR i:=1 TO 7 DO
	IF G.axis[i].Status.Error OR G.power_output[i].Error OR G.reset_output[i].Error THEN
		has_err := TRUE;
		EXIT;
	END_IF
END_FOR

all_powered := TRUE;
FOR i:=1 TO 7 DO
	IF NOT G.power_output[i].Done THEN
		all_powered := FALSE;
		EXIT;
	END_IF
END_FOR

G.estop_hold_req := TRUE;

CASE step OF
0:
	FOR i:=1 TO 7 DO
		G.SetPointGenEnable[i].Execute := FALSE;
		G.SetPointGenDisable[i].Execute := FALSE;
		G.axis_Reset[i].Execute := FALSE;
	END_FOR
	settle_timer(IN:=FALSE);
	step := 1;

1:
	IF has_err THEN
		settle_timer(IN:=FALSE);
		step := 0;
		G.gen_state := _err;
		RETURN;
	END_IF

	IF NOT G.self_check_done THEN
		settle_timer(IN:=FALSE);
		step := 0;
		G.gen_state := _init;
		RETURN;
	END_IF

	IF NOT all_powered THEN
		FOR i:=1 TO 7 DO
			G.power_[i].Enable := TRUE;
		END_FOR
		settle_timer(IN:=FALSE);
		RETURN;
	END_IF

	settle_timer(IN:=TRUE, PT:=T#200MS);
	IF settle_timer.Q THEN
		settle_timer(IN:=FALSE);
		step := 0;
		G.handle_reinit_req := TRUE;
		G.gen_state := _handle;
	END_IF
END_CASE

END_FUNCTION_BLOCK

